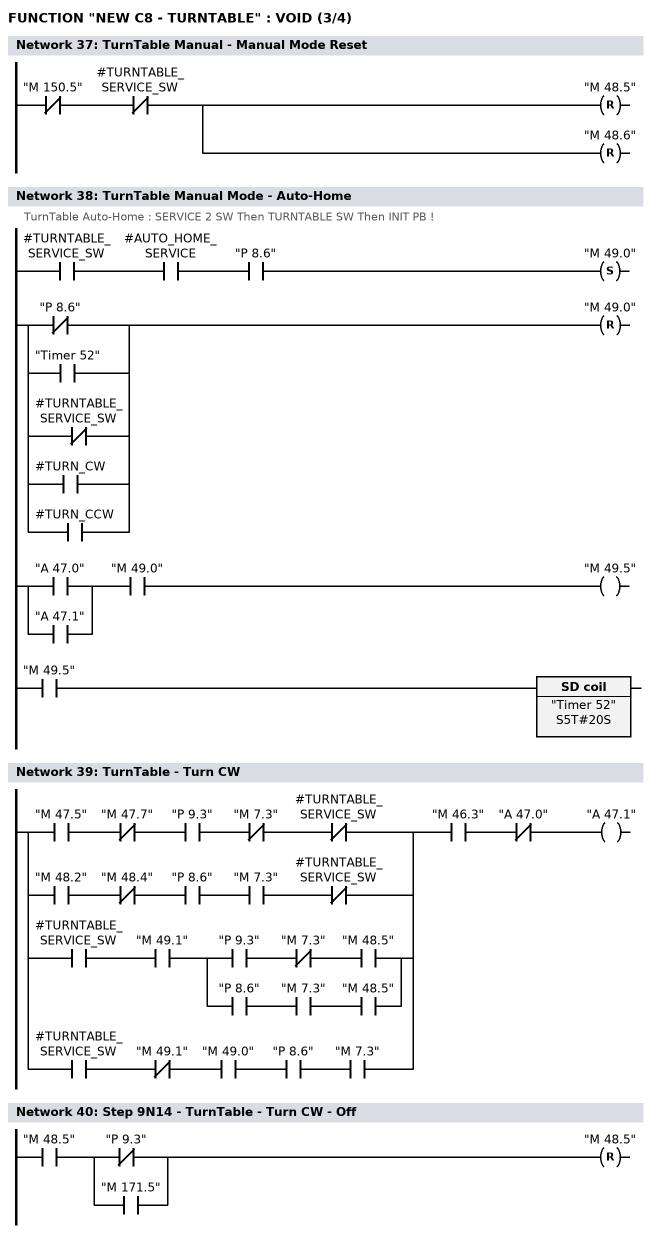

      AN    "M 150.5";
      AN    #TURNTABLE_SERVICE_SW;
      R     "M 48.5";
      R     "M 48.6";
NETWORK
TITLE =TurnTable Manual Mode - Auto-Home
//TurnTable Auto-Home : SERVICE 2 SW Then TURNTABLE SW Then INIT PB !
      A     #TURNTABLE_SERVICE_SW;
      A     #AUTO_HOME_SERVICE;
      A     "P 8.6";
      S     "M 49.0";
//;
      AN    "P 8.6";
      O     "Timer 52";
      ON    #TURNTABLE_SERVICE_SW;
      O     #TURN_CW;
      O     #TURN_CCW;
      R     "M 49.0";
//;
      A(    ;
      O     "A 47.0";
      O     "A 47.1";
      )     ;
      A     "M 49.0";
      =     "M 49.5";
//;
      A     "M 49.5";
      L     S5T#20S;
      SD    "Timer 52";
NETWORK
TITLE =TurnTable - Turn CW

      A(    ;
      A     "M 47.5";
      AN    "M 47.7";
      A     "P 9.3";
      AN    "M 7.3";
      AN    #TURNTABLE_SERVICE_SW;
      O     ;
      A     "M 48.2";
      AN    "M 48.4";
      A     "P 8.6";
      A     "M 7.3";
      AN    #TURNTABLE_SERVICE_SW;
      O     ;
      A     #TURNTABLE_SERVICE_SW;
      A     "M 49.1";
      A(    ;
      A     "P 9.3";
      AN    "M 7.3";
      A     "M 48.5";
      O     ;
      A     "P 8.6";
      A     "M 7.3";
      A     "M 48.5";
      )     ;
      O     ;
      A     #TURNTABLE_SERVICE_SW;
      AN    "M 49.1";
      A     "M 49.0";
      A     "P 8.6";
      A     "M 7.3";
      )     ;
      A     "M 46.3";
      AN    "A 47.0";
      =     "A 47.1";
NETWORK
TITLE =Step 9N14 - TurnTable - Turn CW - Off

      A     "M 48.5";
      A(    ;
      ON    "P 9.3";
      O     "M 171.5";
      )     ;
      R     "M 48.5";
NETWORK
TITLE =Turn Table - Turn CCW
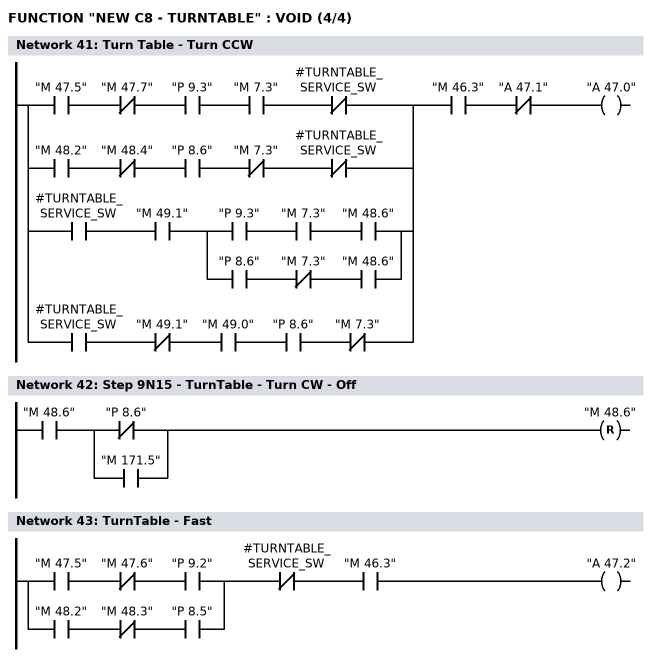

      A(    ;
      A     "M 47.5";
      AN    "M 47.7";
      A     "P 9.3";
      A     "M 7.3";
      AN    #TURNTABLE_SERVICE_SW;
      O     ;
      A     "M 48.2";
      AN    "M 48.4";
      A     "P 8.6";
      AN    "M 7.3";
      AN    #TURNTABLE_SERVICE_SW;
      O     ;
      A     #TURNTABLE_SERVICE_SW;
      A     "M 49.1";
      A(    ;
      A     "P 9.3";
      A     "M 7.3";
      A     "M 48.6";
      O     ;
      A     "P 8.6";
      AN    "M 7.3";
      A     "M 48.6";
      )     ;
      O     ;
      A     #TURNTABLE_SERVICE_SW;
      AN    "M 49.1";
      A     "M 49.0";
      A     "P 8.6";
      AN    "M 7.3";
      )     ;
      A     "M 46.3";
      AN    "A 47.1";
      =     "A 47.0";
NETWORK
TITLE =Step 9N15 - TurnTable - Turn CW - Off

      A     "M 48.6";
      A(    ;
      ON    "P 8.6";
      O     "M 171.5";
      )     ;
      R     "M 48.6";
NETWORK
TITLE =TurnTable - Fast

      A(    ;
      A     "M 47.5";
      AN    "M 47.6";
      A     "P 9.2";
      O     ;
      A     "M 48.2";
      AN    "M 48.3";
      A     "P 8.5";
      )     ;
      AN    #TURNTABLE_SERVICE_SW;
      A     "M 46.3";
      =     "A 47.2";
NETWORK
TITLE =TurnTable Position : Home = DB50.238:1 / Delivery = DB50.238:2

      OPN   "DB LAUER";
      ON    "P 8.6";
      ON    "P 9.3";
      JC    M003;
      L     W#16#0;
      T     DBW  238;
      BEC   ;

M003: A     "P 8.6";
      JC    M004;
      L     W#16#1;
      T     DBW  238;
      BEC   ;

M004: L     W#16#2;
      T     DBW  238;
END_FUNCTION

FUNCTION "NEW C9 - PUSHER 2" : VOID
TITLE =NEW FC950 (was FC1050) - Conveyor 9 / Pusher 2 Pos.11
//
//v1.0 2026-11-24: OMRON HMI positioning time (Timer 62) per packet length class
//from DB15 "PACKET POSITION DB".C9_Stop_S5T (FC1215 "PACKET POSITIONING", called
//by FC942). Class without time = "HMI_DB".CONV_9_POS_mS x 10 as before.
//v1.1 2026-11-24: DB15 symbol renamed "PACKET POSITION DB" - no code change.
NAME : POS_11
VERSION : 1.1


VAR_TEMP
  MAIN_SERVICE_2_SW : BOOL ;
  CONVEYOR_9_RUN : BOOL ;
  PUSHER_PUSH : BOOL ;
  INITIALISATION : BOOL ;
  POSITION_TIME : S5TIME ;
  ZOOLOO : TIME ;
END_VAR
BEGIN
NETWORK
TITLE =Pusher 2 - Service

      A     "HMI_DB".ALL_SERVICE_ENABLE_SW;
      A     "HMI_DB".CONVEYOR_9_SERVICE_SW;
      A     "HMI_DB".SERVICE_SW_2_STATUS;
      =     #MAIN_SERVICE_2_SW;
//;
      A     #MAIN_SERVICE_2_SW;
      O     "M 50.1";
      JNB   CON9;
      A     "HMI_DB".HMI_CONVEYOR_9_TEST_SSW;
      =     #CONVEYOR_9_RUN;
//;
      A     "HMI_DB".HMI_PUSHER_2_TEST_SSW;
      =     #PUSHER_PUSH;
//;
      A     "HMI_DB".SERVICE_INIT_PB;
      =     #INITIALISATION;
//;
      A     #CONVEYOR_9_RUN;
      S     "DB UTILITY".Conveyor_8_Disable;
//;
      A     #PUSHER_PUSH;
      S     "DB UTILITY".Conveyor_9_Disable;
//;
      AN    #MAIN_SERVICE_2_SW;
      R     "HMI_DB".HMI_CONVEYOR_9_TEST_SSW;
      R     "HMI_DB".HMI_PUSHER_2_TEST_SSW;
      R     "DB UTILITY".Conveyor_8_Disable;
      R     "DB UTILITY".Conveyor_9_Disable;

CON9: R     #CONVEYOR_9_RUN;
      R     #PUSHER_PUSH;
      R     #INITIALISATION;
      FP    "FP 169.1";
      =     "M 50.1";
NETWORK
TITLE =Pusher Rollers - Max Run Time

      A     "M 51.2";
      AN    "M 51.3";
      A     "M 0.3";
      L     S5T#5S;
      SD    "Timer 51";
NETWORK
TITLE =Conveyor 9 - Pusher Steps Register - Reset

      A(    ;
      A     "M 52.1";
      O     "Timer 51";
      O     #INITIALISATION;
      O     "DB UTILITY".Conveyor_9_Disable;
      )     ;
      A     "M 0.3";
      JC    M001;
      JU    M002;

M001: L     W#16#0;
      T     "MW 51";
      T     "MB 53";

M002: NOP   0;
NETWORK
TITLE =Step 10N1 - Power ON
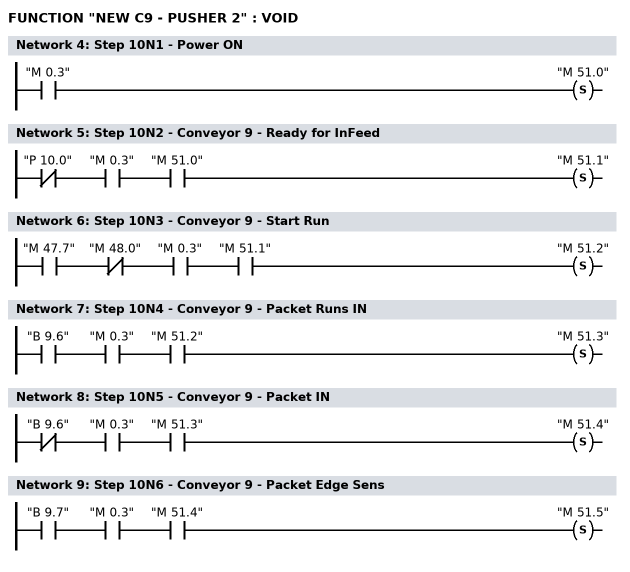

      A     "M 0.3";
      S     "M 51.0";
NETWORK
TITLE =Step 10N2 - Conveyor 9 - Ready for InFeed

      AN    "P 10.0";
      A     "M 0.3";
      A     "M 51.0";
      S     "M 51.1";
NETWORK
TITLE =Step 10N3 - Conveyor 9 - Start Run

      A     "M 47.7";
      AN    "M 48.0";
      A     "M 0.3";
      A     "M 51.1";
      S     "M 51.2";
NETWORK
TITLE =Step 10N4 - Conveyor 9 - Packet Runs IN

      A     "B 9.6";
      A     "M 0.3";
      A     "M 51.2";
      S     "M 51.3";
NETWORK
TITLE =Step 10N5 - Conveyor 9 - Packet IN

      AN    "B 9.6";
      A     "M 0.3";
      A     "M 51.3";
      S     "M 51.4";
NETWORK
TITLE =Step 10N6 - Conveyor 9 - Packet Edge Sens

      A     "B 9.7";
      A     "M 0.3";
      A     "M 51.4";
      S     "M 51.5";
NETWORK
TITLE =Time Convertion - Lateral Packet Position to Feeder - Adj.(HMI)

      A     "M 140.3";
      AN    "M 6.7";
      FP    "FP 147.2";
      JNB   BYP1;
      L     "HMI_DB".CONV_9_POS_mS; // Integer contains MILLISECOND seconds
      L     10;
      *I    ;
      ITD   ;
      T     #ZOOLOO;

      CALL "TIM_S5TI" (
           IN                       := #ZOOLOO,
           RET_VAL                  := #POSITION_TIME);

      L     #POSITION_TIME;
      T     "MW 184";
BYP1: CLR   ;

      A     "M 140.3";
      A     "M 51.5";
      AN    "M 51.6";
      A     "M 0.3";
      L     "PACKET POSITION DB".C9_Stop_S5T; // Was MW 184 - Now per Length Class (DB15)
      SD    "Timer 62"; // OMRON HMI
NETWORK
TITLE =Conveyor 9 - Lateral Packet Position to Feeder - Adj.(HMI)

      AN    "M 140.3";
      AN    "M 6.7";
      FP    "FP 149.5";
      JNB   BYP2;
      OPN   "DB LAUER";
      CALL "LAUER TIME" (
           QUEL                     := DBW  248,
           _TIME                    := MW   124);

BYP2: NOP   0;

      AN    "M 140.3";
      A     "M 51.5";
      AN    "M 51.6";
      A     "M 0.3";
      L     MW   124;
      SD    "Timer 50"; // LAUER HMI
NETWORK
TITLE =Step 10N7 - Conveyor 9 - Packet in Position - Stop
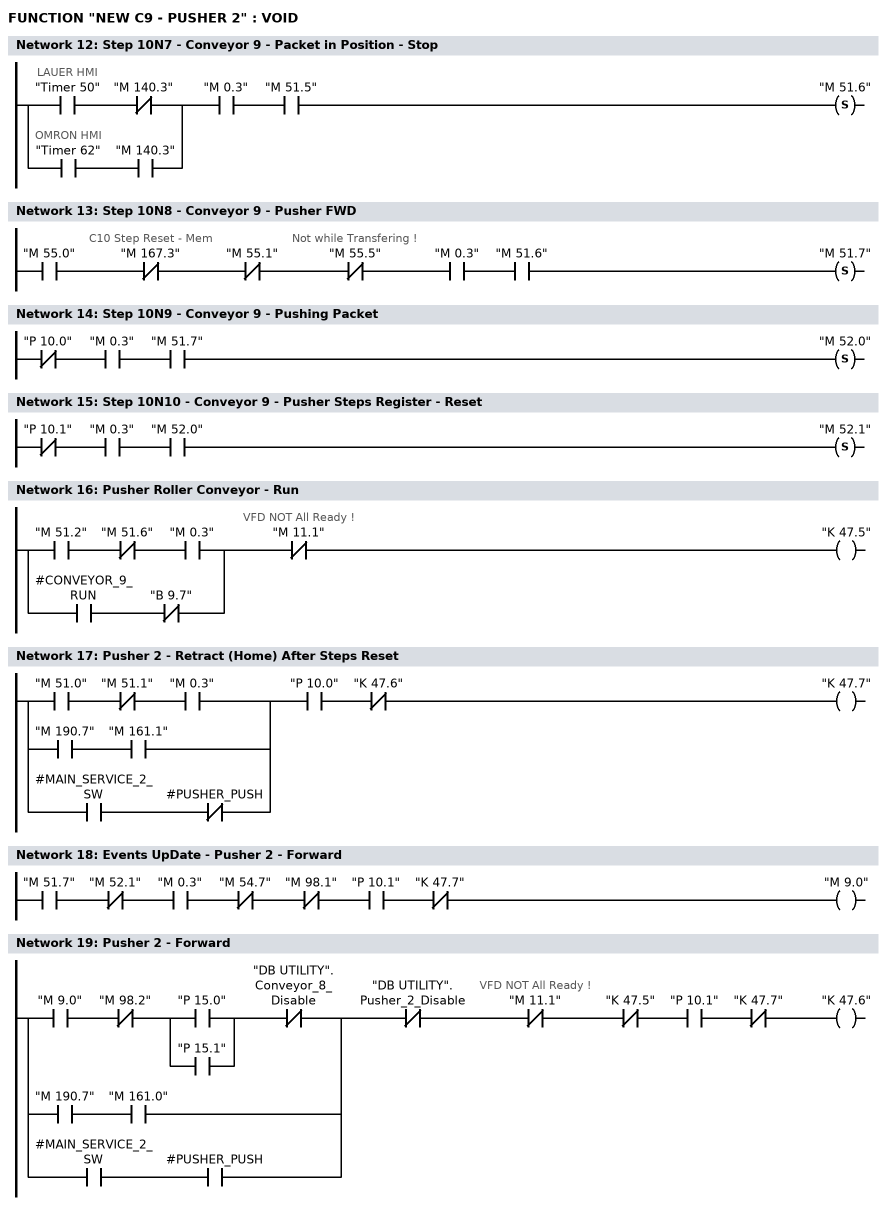

      A(    ;
      O(    ;
      A     "Timer 50"; // LAUER HMI
      AN    "M 140.3";
      )     ;
      O(    ;
      A     "Timer 62"; // OMRON HMI
      A     "M 140.3";
      )     ;
      )     ;
      A     "M 0.3";
      A     "M 51.5";
      S     "M 51.6";
NETWORK
TITLE =Step 10N8 - Conveyor 9 - Pusher FWD

      A     "M 55.0";
      AN    "M 167.3"; // C10 Step Reset - Mem
      AN    "M 55.1";
      AN    "M 55.5"; // Not while Transfering !
      A     "M 0.3";
      A     "M 51.6";
      S     "M 51.7";
NETWORK
TITLE =Step 10N9 - Conveyor 9 - Pushing Packet

      AN    "P 10.0";
      A     "M 0.3";
      A     "M 51.7";
      S     "M 52.0";
NETWORK
TITLE =Step 10N10 - Conveyor 9 - Pusher Steps Register - Reset

      AN    "P 10.1";
      A     "M 0.3";
      A     "M 52.0";
      S     "M 52.1";
NETWORK
TITLE =Pusher Roller Conveyor - Run

      A     "M 51.2";
      AN    "M 51.6";
      A     "M 0.3";
      O(    ;
      A     #CONVEYOR_9_RUN;
      AN    "B 9.7";
      )     ;
      AN    "M 11.1"; // VFD NOT All Ready !
      =     "K 47.5";
NETWORK
TITLE =Pusher 2 - Retract (Home) After Steps Reset

      A(    ;
      A     "M 51.0";
      AN    "M 51.1";
      A     "M 0.3";
      O     ;
      A     "M 190.7";
      A     "M 161.1";
      O     ;
      A     #MAIN_SERVICE_2_SW;
      AN    #PUSHER_PUSH;
      )     ;
      A     "P 10.0";
      AN    "K 47.6";
      =     "K 47.7";
NETWORK
TITLE =Events UpDate - Pusher 2 - Forward

      A     "M 51.7";
      AN    "M 52.1";
      A     "M 0.3";
      AN    "M 54.7";
      AN    "M 98.1";
      A     "P 10.1";
      AN    "K 47.7";
      =     "M 9.0";
NETWORK
TITLE =Pusher 2 - Forward

      A(    ;
      A     "M 9.0";
      AN    "M 98.2";
      A(    ;
      O     "P 15.0";
      O     "P 15.1";
      )     ;
      AN    "DB UTILITY".Conveyor_8_Disable;
      O     ;
      A     "M 190.7";
      A     "M 161.0";
      O     ;
      A     #MAIN_SERVICE_2_SW;
      A     #PUSHER_PUSH;
      )     ;
      AN    "DB UTILITY".Pusher_2_Disable;
      AN    "M 11.1"; // VFD NOT All Ready !
      AN    "K 47.5";
      A     "P 10.1";
      AN    "K 47.7";
      =     "K 47.6";
NETWORK
TITLE =Position Data Return

      OPN   "DB LAUER";
//;
      ON    "P 10.0";
      ON    "P 10.1";
      JC    M003;
      L     W#16#0;
      T     DBW  220;
      BEC   ;

M003: AN    "P 10.0";
      JC    M004;
      L     W#16#1;
      T     DBW  220;
      BEC   ;

M004: L     W#16#2;
      T     DBW  220;
END_FUNCTION

FUNCTION "NEW C10 - PIVOT PIW" : VOID
TITLE =FC 955 > NEW FC954 (was FC1054) - Pivot Conveyor 10 - Collator
//v0.1 2026-11-19: C10 encoder Ch5 read DIRECT every scan: PIW 334 (HW Config)
//instead
//of ACT_CNTV5. Ch4 (width gate) stays ACT_CNTV4: not in the direct area.
NAME : POS_12
VERSION : 0.1


VAR_TEMP
  MAIN_SERVICE_2_SW : BOOL ;
  PIVOT_SERVICE_SW : BOOL ;
  PIVOT_UP : BOOL ;
  PIVOT_DN : BOOL ;
  CONVEYOR_RUN : BOOL ;
  INITIALISATION : BOOL ;
  BARRIER_BLINKER : BOOL ;	//Feeder Safety Light Barrier
  PACKET_WIDTH_10 : WORD ;	//Collator Conveyor 10 - Packet Width
  FRAC_PACKET_WIDTH_10 : WORD ;	//Collator Conveyor 10 - Fraction of Packet Width
  PACKET_WIDTH_FRAC_10 : WORD ;	//Collator Conveyor 10 - Packet Width + Fraction
  SURFACE_LENGTH_LEFT_10 : WORD ;	//Collator Conveyor 10 - Surface Length Left
  QTY_MAX_10 : REAL ;
END_VAR
BEGIN
NETWORK
TITLE =Pivot Service

      A     "HMI_DB".ALL_SERVICE_ENABLE_SW;
      A     "HMI_DB".CONVEYOR_10_SERVICE_SW;
      A     "HMI_DB".SERVICE_SW_2_STATUS;
      =     #MAIN_SERVICE_2_SW;
//;
      A     #MAIN_SERVICE_2_SW;
      O     "M 54.3";
      JNB   PIVO;

      A     "HMI_DB".HMI_PIVOT_SERVICE_SSW;
      =     #PIVOT_SERVICE_SW;
      R     "HMI_DB".HMI_CONVEYOR_10_TEST_SSW;
//;
      A     "HMI_DB".HMI_CONVEYOR_10_TEST_SSW;
      =     #CONVEYOR_RUN;
      R     "HMI_DB".HMI_PIVOT_SERVICE_SSW;
//;
      A(    ;
      O     #PIVOT_SERVICE_SW;
      O     #CONVEYOR_RUN;
      )     ;
      S     "DB UTILITY".Pusher_2_Disable;
//;
      A     #PIVOT_SERVICE_SW;
      A     "HMI_DB".HMI_PIVOT_TEST_DN_SSW;
      AN    "HMI_DB".HMI_PIVOT_TEST_UP_SSW; // Not Both Switches
      =     #PIVOT_DN;
//;
      A     #PIVOT_SERVICE_SW;
      A     "HMI_DB".HMI_PIVOT_TEST_UP_SSW;
      AN    "HMI_DB".HMI_PIVOT_TEST_DN_SSW; // Not Both Switches
      =     #PIVOT_UP;
//;
      AN(   ;
      O     "P 15.0";
      O     "P 15.1";
      )     ;
      R     #CONVEYOR_RUN;
//;
      A     "HMI_DB".SERVICE_INIT_PB;
      =     #INITIALISATION;
//;
      AN    #MAIN_SERVICE_2_SW;
      R     "HMI_DB".HMI_PIVOT_SERVICE_SSW;
      R     "HMI_DB".HMI_CONVEYOR_10_TEST_SSW;
      R     "HMI_DB".HMI_PIVOT_TEST_DN_SSW;
      R     "HMI_DB".HMI_PIVOT_TEST_UP_SSW;
      R     "DB UTILITY".Pusher_2_Disable;

PIVO: R     #PIVOT_SERVICE_SW;
      R     #CONVEYOR_RUN;
      R     #INITIALISATION;
      R     #PIVOT_DN;
      R     #PIVOT_UP;
      FP    "FP 169.2";
      =     "M 54.3";
NETWORK
TITLE =Conveyor 10 - Packet Width - Measurements [mS]

      A     "B 10.4"; // C10 InFeed Sens
      A     "M 55.1"; // Collator Trigger - Step
      S     "M 166.4";
//;
      A     "M 166.4";
      =     "FM350 DB".CONTROL_SIGNALS.SW_GATE4;
//;
      A     "M 166.4";
      FP    "FP 149.7";
      JNB   NRAZ;
      L     0;
      T     "COLLATORS DB".Packet_Width_C10_mS;

NRAZ: A     "M 166.4";
      JNB   NCNT;
      L     "COLLATORS DB".Packet_Width_C10_mS;
      L     "DB UTILITY".Scan_Cycle_Previous;
      ITD   ;
      +D    ;
      T     "COLLATORS DB".Packet_Width_C10_mS;

NCNT: A     "M 166.4";
      AN    "B 10.4";
      JNB   M104;
      L     "FM350 DB".ACT_CNTV4; // C10 Encoder Counter
      T     #PACKET_WIDTH_10;
      T     "COLLATORS DB".Packet_Width_C10;
//;
      L     #PACKET_WIDTH_10;
      ITD   ;
      DTR   ;
      L     2.000000e-001;
      *R    ;
      RND   ;

      T     "COLLATORS DB".Frac_Packet_Width_C10;

      T     #FRAC_PACKET_WIDTH_10;
      L     #PACKET_WIDTH_10;
      +I    ;
      T     "COLLATORS DB".Packet_Width_Frac_C10;
      T     #PACKET_WIDTH_FRAC_10;
      R     "M 166.4";
      S     "M 167.2";

M104: NOP   0;
NETWORK
TITLE =Conveyor 10 - Packet Width Measurements [mm] - While Collating

      A     "B 10.4"; // C10 InFeed Sens - New Packet
      FP    "M 188.5";
      A     "A 48.0";
      JCN   NPRT;

      L     "PIW 334"; // Direct Ch5 (was ACT_CNTV5, ~100 mS old) C10 Encoder Counter
      T     "HOUSE_KEEPING DB".C10_Encoder_READ_Mem;

NPRT: AN    "B 10.4"; // C10 InFeed Sens - New Packet End
      FP    "M 188.6";
      JCN   NTKE;

      L     "PIW 334"; // Direct Ch5 (was ACT_CNTV5, ~100 mS old) C10 Encoder Counter
      L     "HOUSE_KEEPING DB".C10_Encoder_READ_Mem;
      -I    ;
      T     "HOUSE_KEEPING DB".C10_Packet_Width_ep; // C4 Packet Length [ep]
      DTR   ;
//;
      L     3.100000e-001; //  Encoder Wheel 283mm / 600 PPR  [mm/pulse]
      *R    ;
      RND   ;
      T     "HOUSE_KEEPING DB".C10_Packet_Width_mm;

NTKE: NOP   0;
NETWORK
TITLE =Conveyor 10 - Packet Width Measurements [mS]
//Conveyor 10 - Packet Width Measurements [mS]


NETWORK
TITLE =Conveyor 10 - Surface Length Left (PulseUnit) - Measurements

      A     "M 166.5";
      =     "FM350 DB".CONTROL_SIGNALS.SW_GATE5;
//;
      A     "M 166.5";
      JNB   M665;
      L     "COLLATORS DB".Surface_Length_10;
      L     "PIW 334"; // Direct Ch5 (was ACT_CNTV5, ~100 mS old)
      -D    ;
      T     #SURFACE_LENGTH_LEFT_10;
      L     0;
      >=I   ;
      JNB   T010;
      L     #SURFACE_LENGTH_LEFT_10;
      T     "COLLATORS DB".Surface_Length_Left_10;

T010: NOP   0;

M665: NOP   0;

      A     "M 55.1"; // Collator Trigger
      FP    "FP 154.6";
      S     "M 166.5";
NETWORK
TITLE =Conveyor 10 - Space Between Packet - Calculator
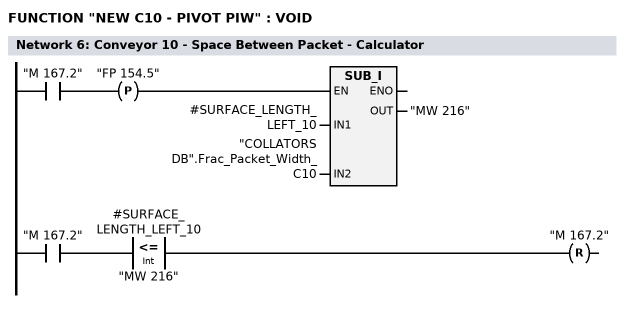

      A     "M 167.2";
      FP    "FP 154.5";
      JNB   M582;
      L     #SURFACE_LENGTH_LEFT_10;
      L     "COLLATORS DB".Frac_Packet_Width_C10;
      -I    ;
      T     "MW 216";

M582: NOP   0;

      A     "M 167.2";
      A(    ;
      L     #SURFACE_LENGTH_LEFT_10;
      L     "MW 216";
      <=I   ;
      )     ;
      R     "M 167.2";
NETWORK
TITLE =Conveyor 10 - Collating Surface Manager

      A     "M 166.5";
      AN    "M 55.4";
      AN    "M 54.4"; // Collator Full - Count Flag Off
      A     "M 55.3";
      JNB   M554;

      A(    ;
      L     #SURFACE_LENGTH_LEFT_10;
      L     "COLLATORS DB".Packet_Width_Frac_C10;
      <I    ;
      )     ;
      S     "M 54.4"; // Collator Full - Count - Set

M554: NOP   0;

      A     "M 167.3"; // C10 Step Reset - Mem
      R     "M 54.4"; // Collator Full - Count - Reset
NETWORK
TITLE =Conveyor 10 - Surface Length Reset

      ON(   ;
      O     "P 15.0"; // While C10 Pivoting...
      O     "P 15.1";
      )     ;
      L     S5T#200MS;
      SD    "Timer 104";
//;
      A     "Timer 104"; // C10 Surface Length Reset
      R     "M 166.4";
      R     "M 166.5";
NETWORK
TITLE =Clearing - C10 Counters Reset
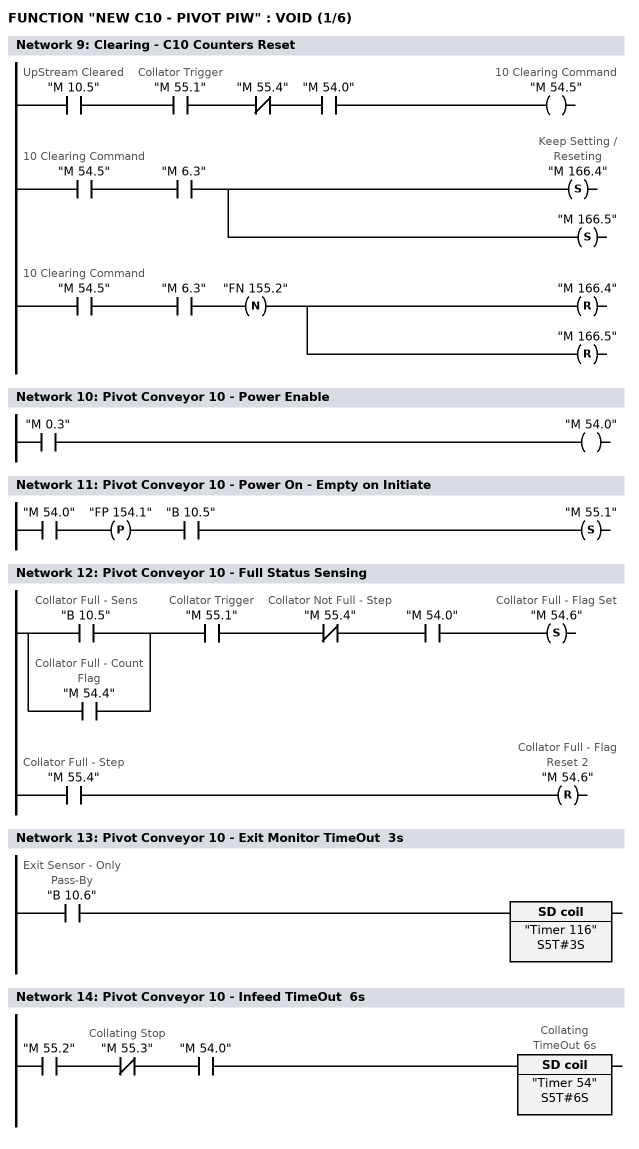

      A     "M 10.5"; // UpStream Cleared
      A     "M 55.1"; // Collator Trigger
      AN    "M 55.4";
      A     "M 54.0";
      =     "M 54.5"; // 10 Clearing Command
//;
      A     "M 54.5"; // 10 Clearing Command
      A     "M 6.3";
      S     "M 166.4"; // Keep Setting / Reseting
      S     "M 166.5";
//;
      A     "M 54.5"; // 10 Clearing Command
      A     "M 6.3";
      FN    "FN 155.2";
      R     "M 166.4";
      R     "M 166.5";
NETWORK
TITLE =Pivot Conveyor 10 - Power Enable

      A     "M 0.3";
      =     "M 54.0";
NETWORK
TITLE =Pivot Conveyor 10 - Power On - Empty on Initiate

      A     "M 54.0";
      FP    "FP 154.1"; // Empty on Power ON
      A     "B 10.5";
      S     "M 55.1";
NETWORK
TITLE =Pivot Conveyor 10 - Full Status Sensing

      A(    ;
      O     "B 10.5"; // Collator Full - Sens
      O     "M 54.4"; // Collator Full - Count Flag
      )     ;
      A     "M 55.1"; // Collator Trigger
      AN    "M 55.4"; // Collator Not Full - Step
      A     "M 54.0";
      S     "M 54.6"; // Collator Full - Flag Set
//;
      A     "M 55.4"; // Collator Full - Step
      R     "M 54.6"; // Collator Full - Flag Reset 2
NETWORK
TITLE =Pivot Conveyor 10 - Exit Monitor TimeOut  3s

      A     "B 10.6"; // Exit Sensor - Only Pass-By
      L     S5T#3S;
      SD    "Timer 116"; // Packet is Stuck !
NETWORK
TITLE =Pivot Conveyor 10 - Infeed TimeOut  6s

      A     "M 55.2";
      AN    "M 55.3"; // Collating Stop
      A     "M 54.0";
      L     S5T#6S; // Collating TimeOut 6s
      SD    "Timer 54";
NETWORK
TITLE =Pivot Conveyor 10 - Fault
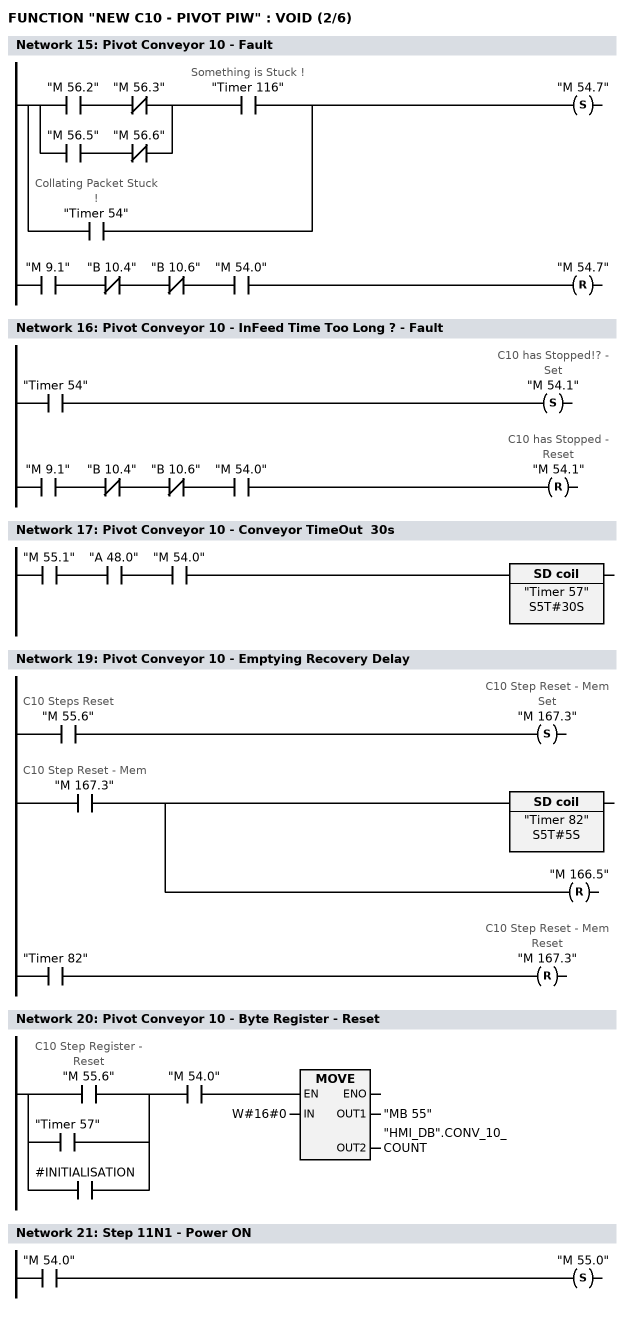

      A(    ;
      A(    ;
      A     "M 56.2";
      AN    "M 56.3";
      O     ;
      A     "M 56.5";
      AN    "M 56.6";
      )     ;
      A     "Timer 116"; // Something is Stuck !
      O     "Timer 54"; // Collating Packet Stuck !
      )     ;
      S     "M 54.7";
//;
      A     "M 9.1";
      AN    "B 10.4";
      AN    "B 10.6";
      A     "M 54.0";
      R     "M 54.7";
NETWORK
TITLE =Pivot Conveyor 10 - InFeed Time Too Long ? - Fault

      A     "Timer 54";
      S     "M 54.1"; // C10 has Stopped!? - Set
//;
      A     "M 9.1";
      AN    "B 10.4";
      AN    "B 10.6";
      A     "M 54.0";
      R     "M 54.1"; // C10 has Stopped - Reset
NETWORK
TITLE =Pivot Conveyor 10 - Conveyor TimeOut  30s

      A     "M 55.1";
      A     "A 48.0";
      A     "M 54.0";
      L     S5T#30S;
      SD    "Timer 57";
NETWORK
TITLE =Collating
//Collating


NETWORK
TITLE =Pivot Conveyor 10 - Emptying Recovery Delay

      A     "M 55.6"; // C10 Steps Reset
      S     "M 167.3"; // C10 Step Reset - Mem Set
//;
      A     "M 167.3"; // C10 Step Reset - Mem
      L     S5T#5S;
      SD    "Timer 82";
      R     "M 166.5";
//;
      A     "Timer 82";
      R     "M 167.3"; // C10 Step Reset - Mem Reset
NETWORK
TITLE =Pivot Conveyor 10 - Byte Register - Reset

      A(    ;
      O     "M 55.6"; // C10 Step Register - Reset
      O     "Timer 57";
      O     #INITIALISATION;
      )     ;
      A     "M 54.0";
      JNB   M001;
      L     W#16#0;
      T     "MB 55";
      T     "HMI_DB".CONV_10_COUNT;

M001: NOP   0;
NETWORK
TITLE =Step 11N1 - Power ON

      A     "M 54.0";
      S     "M 55.0";
NETWORK
TITLE =Step 11N2 - Conveyor 10 - Run
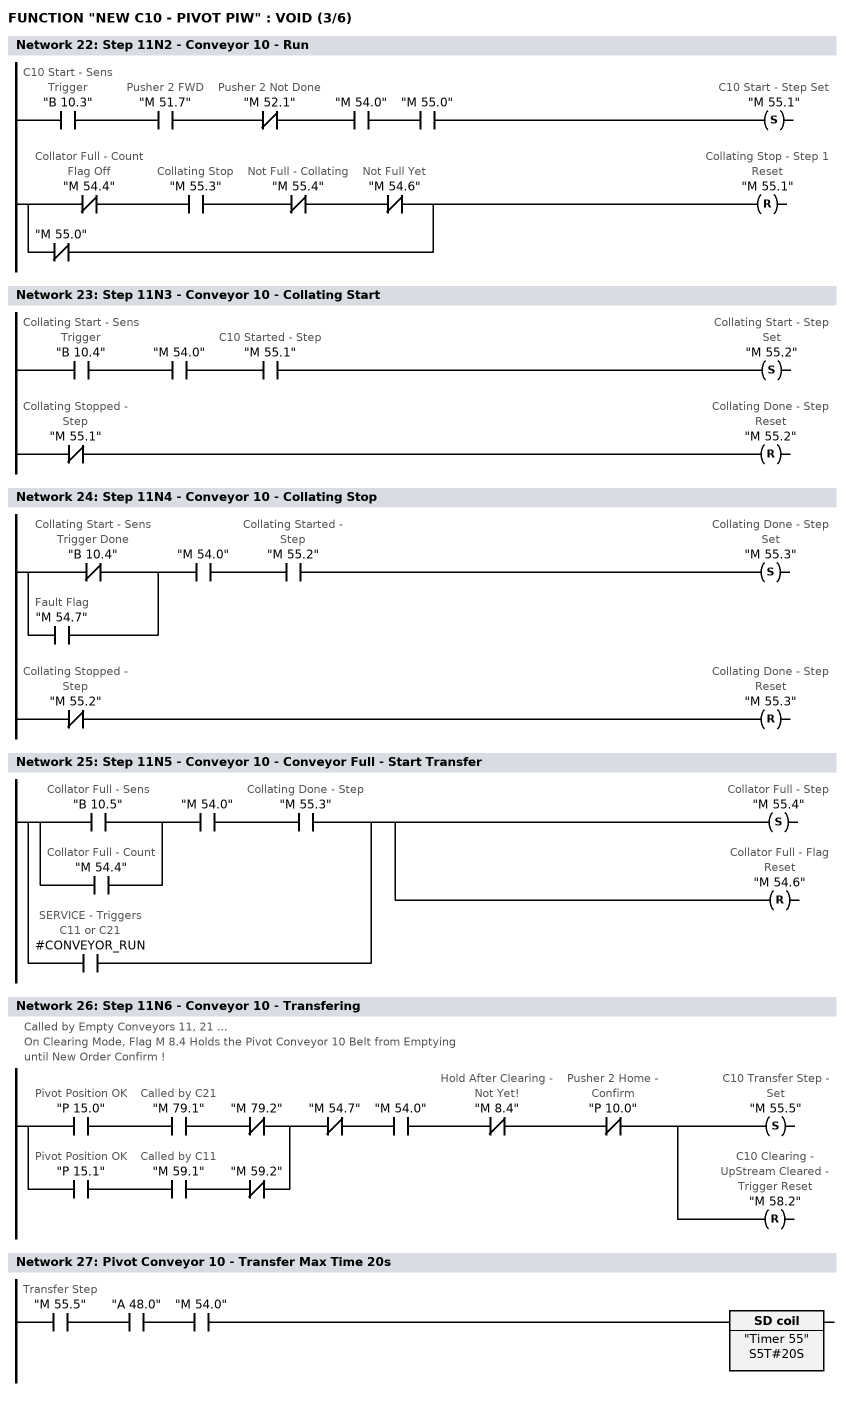

      A     "B 10.3"; // C10 Start - Sens Trigger
      A     "M 51.7"; // Pusher 2 FWD
      AN    "M 52.1"; // Pusher 2 Not Done
      A     "M 54.0";
      A     "M 55.0";
      S     "M 55.1"; // C10 Start - Step Set
//;
      A(    ;
      AN    "M 54.4"; // Collator Full - Count Flag Off
      A     "M 55.3"; // Collating Stop
      AN    "M 55.4"; // Not Full - Collating
      AN    "M 54.6"; // Not Full Yet
      ON    "M 55.0";
      )     ;
      R     "M 55.1"; // Collating Stop - Step 1 Reset
NETWORK
TITLE =Step 11N3 - Conveyor 10 - Collating Start

      A     "B 10.4"; // Collating Start - Sens Trigger
      A     "M 54.0";
      A     "M 55.1"; // C10 Started - Step
      S     "M 55.2"; // Collating Start - Step Set
//;
      AN    "M 55.1"; // Collating Stopped - Step
      R     "M 55.2"; // Collating Done - Step Reset
NETWORK
TITLE =Step 11N4 - Conveyor 10 - Collating Stop

      A(    ;
      ON    "B 10.4"; // Collating Start - Sens Trigger Done
      O     "M 54.7"; // Fault Flag
      )     ;
      A     "M 54.0";
      A     "M 55.2"; // Collating Started - Step
      S     "M 55.3"; // Collating Done - Step Set
//;
      AN    "M 55.2"; // Collating Stopped - Step
      R     "M 55.3"; // Collating Done - Step Reset
NETWORK
TITLE =Step 11N5 - Conveyor 10 - Conveyor Full - Start Transfer

      A(    ;
      O     "B 10.5"; // Collator Full - Sens
      O     "M 54.4"; // Collator Full - Count
      )     ;
      A     "M 54.0";
      A     "M 55.3"; // Collating Done - Step
      O     #CONVEYOR_RUN; // SERVICE - Triggers C11 or C21
      S     "M 55.4"; // Collator Full - Step
      R     "M 54.6"; // Collator Full - Flag Reset
NETWORK
TITLE =Step 11N6 - Conveyor 10 - Transfering
//Called by Empty Conveyors 11, 21 ...
//On Clearing Mode, Flag M 8.4 Holds the Pivot Conveyor 10 Belt from Emptying
//until New Order Confirm !
      A(    ;
      A     "P 15.0"; // Pivot Position OK
      A     "M 79.1"; // Called by C21
      AN    "M 79.2";
      O     ;
      A     "P 15.1"; // Pivot Position OK
      A     "M 59.1"; // Called by C11
      AN    "M 59.2";
      )     ;
      AN    "M 54.7";
      A     "M 54.0";
      AN    "M 8.4"; // Hold After Clearing - Not Yet!
      AN    "P 10.0"; // Pusher 2 Home - Confirm
      S     "M 55.5"; // C10 Transfer Step - Set
      R     "M 58.2"; // C10 Clearing - UpStream Cleared - Trigger Reset
NETWORK
TITLE =Pivot Conveyor 10 - Transfer Max Time 20s

      A     "M 55.5"; // Transfer Step
      A     "A 48.0";
      A     "M 54.0";
      L     S5T#20S;
      SD    "Timer 55"; // Transfer TimeOut
NETWORK
TITLE =Step 11N7 - Conveyor 10 - Steps Register - Reset
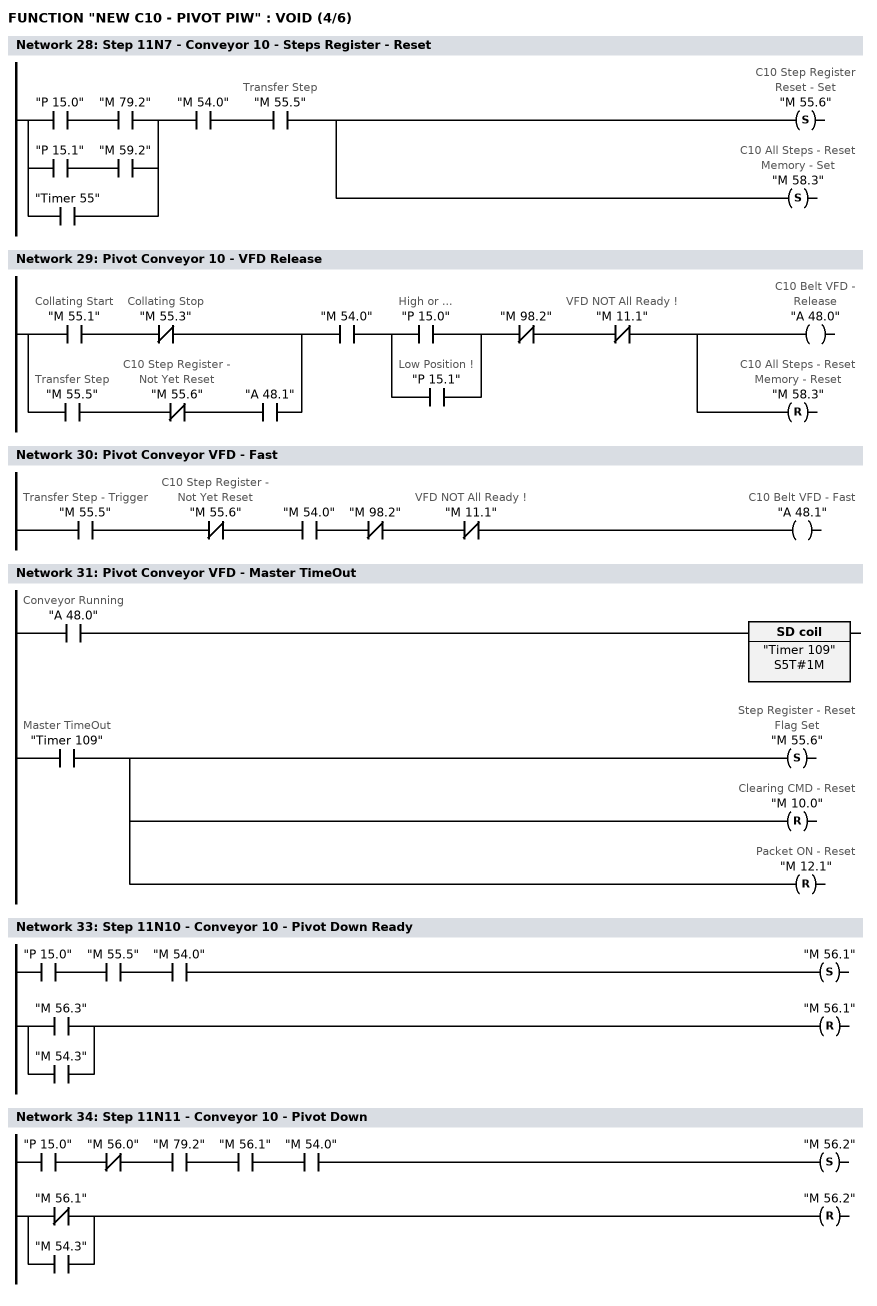

      A(    ;
      A     "P 15.0";
      A     "M 79.2";
      O     ;
      A     "P 15.1";
      A     "M 59.2";
      O     "Timer 55";
      )     ;
      A     "M 54.0";
      A     "M 55.5"; // Transfer Step
      S     "M 55.6"; // C10 Step Register Reset - Set
      S     "M 58.3"; // C10 All Steps - Reset Memory - Set
NETWORK
TITLE =Pivot Conveyor 10 - VFD Release

      A(    ;
      A     "M 55.1"; // Collating Start
      AN    "M 55.3"; // Collating Stop
      O     ;
      A     "M 55.5"; // Transfer Step
      AN    "M 55.6"; // C10 Step Register - Not Yet Reset
      A     "A 48.1";
      )     ;
      A     "M 54.0";
      A(    ;
      O     "P 15.0"; // High or ...
      O     "P 15.1"; // Low Position !
      )     ;
      AN    "M 98.2";
      AN    "M 11.1"; // VFD NOT All Ready !
      =     "A 48.0"; // C10 Belt VFD - Release
      R     "M 58.3"; // C10 All Steps - Reset Memory - Reset
NETWORK
TITLE =Pivot Conveyor VFD - Fast

      A     "M 55.5"; // Transfer Step - Trigger
      AN    "M 55.6"; // C10 Step Register - Not Yet Reset
      A     "M 54.0";
      AN    "M 98.2";
      AN    "M 11.1"; // VFD NOT All Ready !
      =     "A 48.1"; // C10 Belt VFD - Fast
NETWORK
TITLE =Pivot Conveyor VFD - Master TimeOut

      A     "A 48.0"; // Conveyor Running
      L     S5T#1M;
      SD    "Timer 109"; // Master TimeOut
//;
      A     "Timer 109"; // Master TimeOut
      S     "M 55.6"; // Step Register - Reset Flag Set
      R     "M 10.0"; // Clearing CMD - Reset
      R     "M 12.1"; // Packet ON - Reset
NETWORK
TITLE =Pivot Action
//Pivot Action


NETWORK
TITLE =Step 11N10 - Conveyor 10 - Pivot Down Ready

      A     "P 15.0";
      A     "M 55.5";
      A     "M 54.0";
      S     "M 56.1";
//;
      A     "M 56.3";
      O     "M 54.3";
      R     "M 56.1";
NETWORK
TITLE =Step 11N11 - Conveyor 10 - Pivot Down

      A     "P 15.0";
      AN    "M 56.0";
      A     "M 79.2";
      A     "M 56.1";
      A     "M 54.0";
      S     "M 56.2";
//;
      AN    "M 56.1";
      O     "M 54.3";
      R     "M 56.2";
NETWORK
TITLE =Step 11N12 - Conveyor 10 - Move Dn Stop
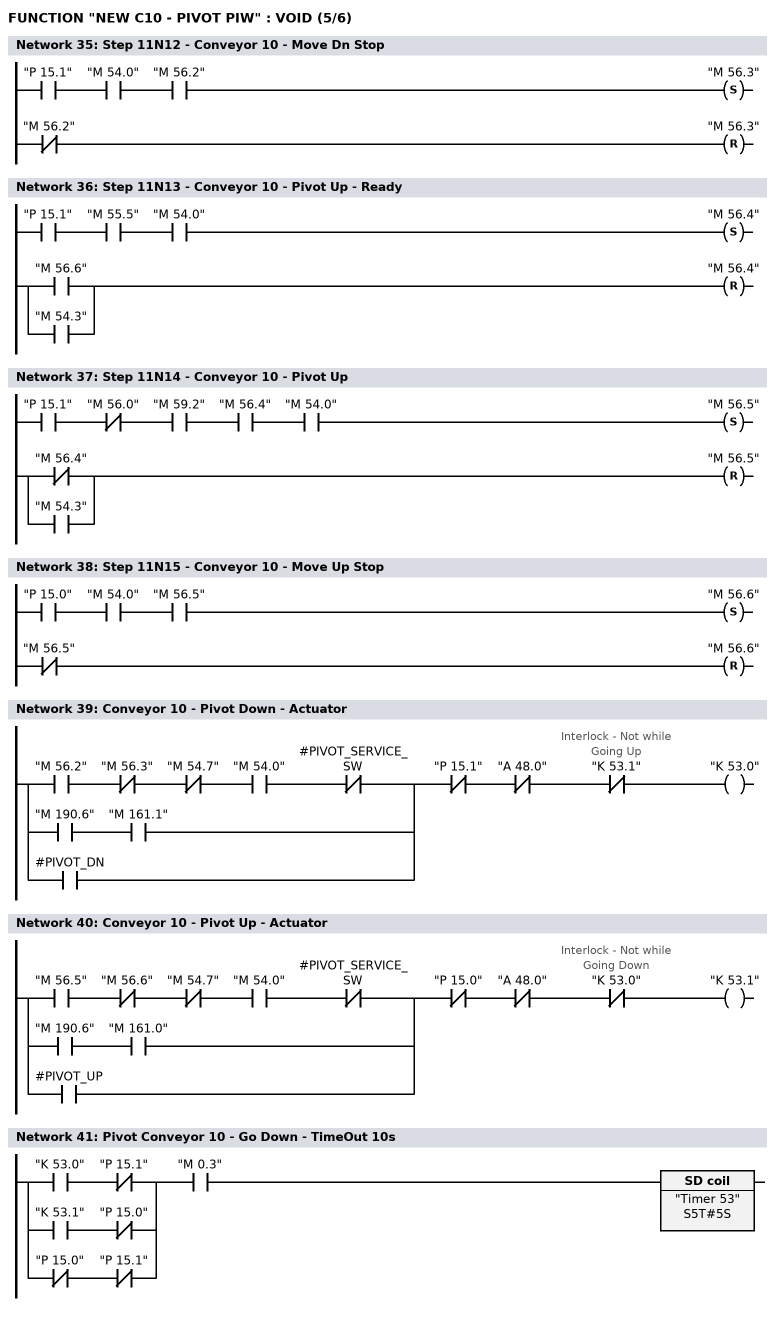

      A     "P 15.1";
      A     "M 54.0";
      A     "M 56.2";
      S     "M 56.3";
//;
      AN    "M 56.2";
      R     "M 56.3";
NETWORK
TITLE =Step 11N13 - Conveyor 10 - Pivot Up - Ready

      A     "P 15.1";
      A     "M 55.5";
      A     "M 54.0";
      S     "M 56.4";
//;
      A     "M 56.6";
      O     "M 54.3";
      R     "M 56.4";
NETWORK
TITLE =Step 11N14 - Conveyor 10 - Pivot Up

      A     "P 15.1";
      AN    "M 56.0";
      A     "M 59.2";
      A     "M 56.4";
      A     "M 54.0";
      S     "M 56.5";
//;
      AN    "M 56.4";
      O     "M 54.3";
      R     "M 56.5";
NETWORK
TITLE =Step 11N15 - Conveyor 10 - Move Up Stop

      A     "P 15.0";
      A     "M 54.0";
      A     "M 56.5";
      S     "M 56.6";
//;
      AN    "M 56.5";
      R     "M 56.6";
NETWORK
TITLE =Conveyor 10 - Pivot Down - Actuator

      A(    ;
      A     "M 56.2";
      AN    "M 56.3";
      AN    "M 54.7";
      A     "M 54.0";
      AN    #PIVOT_SERVICE_SW;
      O     ;
      A     "M 190.6";
      A     "M 161.1";
      )     ;
      O     #PIVOT_DN;
      AN    "P 15.1";
      AN    "A 48.0";
      AN    "K 53.1"; // Interlock - Not while Going Up
      =     "K 53.0";
NETWORK
TITLE =Conveyor 10 - Pivot Up - Actuator

      A(    ;
      A     "M 56.5";
      AN    "M 56.6";
      AN    "M 54.7";
      A     "M 54.0";
      AN    #PIVOT_SERVICE_SW;
      O     ;
      A     "M 190.6";
      A     "M 161.0";
      )     ;
      O     #PIVOT_UP;
      AN    "P 15.0";
      AN    "A 48.0";
      AN    "K 53.0"; // Interlock - Not while Going Down
      =     "K 53.1";
NETWORK
TITLE =Pivot Conveyor 10 - Go Down - TimeOut 10s

      A(    ;
      A     "K 53.0";
      AN    "P 15.1";
      O     ;
      A     "K 53.1";
      AN    "P 15.0";
      O     ;
      AN    "P 15.0";
      AN    "P 15.1";
      )     ;
      A     "M 0.3";
      L     S5T#5S;
      SD    "Timer 53";
NETWORK
TITLE =Pivot Conveyor 10 - Pivot Alarm
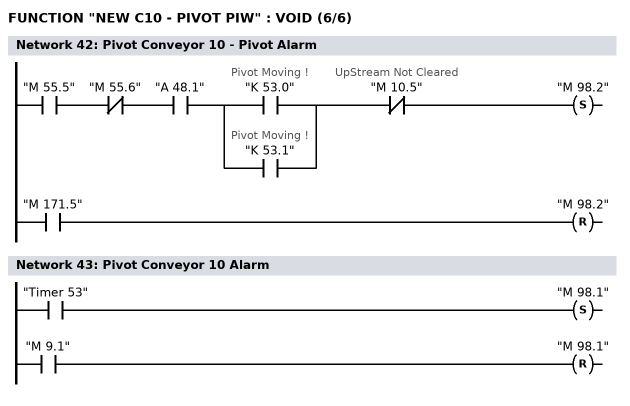

      A(    ;
      A     "M 55.5";
      AN    "M 55.6";
      A     "A 48.1";
      )     ;
      A(    ;
      O     "K 53.0"; // Pivot Moving !
      O     "K 53.1"; // Pivot Moving !
      )     ;
      AN    "M 10.5"; // UpStream Not Cleared
      S     "M 98.2";
//;
      A     "M 171.5";
      R     "M 98.2";
NETWORK
TITLE =Pivot Conveyor 10 Alarm

      A     "Timer 53";
      S     "M 98.1";
//;
      A     "M 9.1";
      R     "M 98.1";
NETWORK
TITLE =DBW  236 - Conveyor 10 - Position Transfer

      OPN   "DB LAUER";

      O     "P 15.0";
      O     "P 15.1";
      JC    M003;
      L     W#16#0;
      T     DBW  236;
      BEC   ;

M003: AN    "P 15.1";
      JC    M004;
      L     W#16#1;
      T     DBW  236;
      BEC   ;

M004: L     W#16#2;
      T     DBW  236;
END_FUNCTION

FUNCTION "NEW C11 - LINK 1 LO" : VOID
TITLE =NEW FC958 (was FC1058) - Conveyor 11 - Link 1L Pos. 13 Low Level
//
//v0.1 2026-11-19: clearing trigger M9.3 only if pivot LOW (P15.1).
NAME : POS_13_L
VERSION : 0.1


VAR_TEMP
  MAIN_SERVICE_2_SW : BOOL ;
  SERVICE_RUN : BOOL ;
  INITIALISATION : BOOL ;
  BARRIER_BLINKER : BOOL ;
END_VAR
BEGIN
NETWORK
TITLE =Conveyor 11 - Service

      A     "HMI_DB".ALL_SERVICE_ENABLE_SW;
      A     "HMI_DB".CONVEYOR_11_SERVICE_SW;
      A     "HMI_DB".SERVICE_SW_2_STATUS;
      =     #MAIN_SERVICE_2_SW;
//;
      A     #MAIN_SERVICE_2_SW;
      O     "M 58.7";
      JNB   CO11;
//;
      A     "HMI_DB".HMI_CONVEYOR_11_TEST_SSW;
      AN    "A 48.0";
      =     #SERVICE_RUN;
      S     "DB UTILITY".Conveyor_10_Disable;
      S     "DB UTILITY".Pivot_Disable;
//;
      A     "HMI_DB".SERVICE_INIT_PB;
      =     #INITIALISATION;
//;
      AN    #MAIN_SERVICE_2_SW;
      R     "HMI_DB".HMI_CONVEYOR_11_TEST_SSW;
      R     "DB UTILITY".Conveyor_10_Disable;
      R     "DB UTILITY".Pivot_Disable;

CO11: R     #SERVICE_RUN;
      R     #INITIALISATION;
      FP    "FP 148.0";
      =     "M 58.7";
NETWORK
TITLE =Power Enable
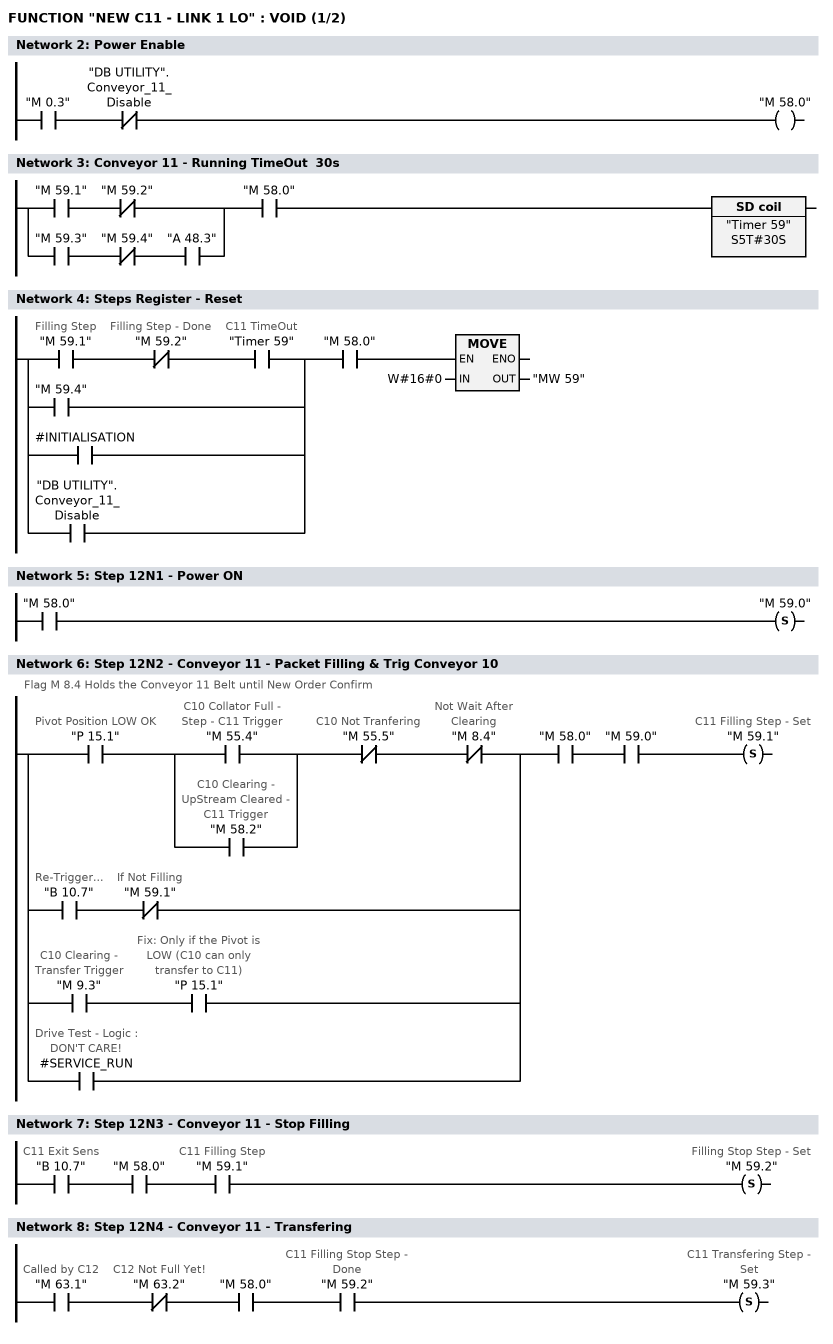

      A     "M 0.3";
      AN    "DB UTILITY".Conveyor_11_Disable;
      =     "M 58.0";
NETWORK
TITLE =Conveyor 11 - Running TimeOut  30s

      A(    ;
      A     "M 59.1";
      AN    "M 59.2";
      O     ;
      A     "M 59.3";
      AN    "M 59.4";
      A     "A 48.3";
      )     ;
      A     "M 58.0";
      L     S5T#30S;
      SD    "Timer 59"; // C11 TimeOut
NETWORK
TITLE =Steps Register - Reset

      A(    ;
      A     "M 59.1"; // Filling Step
      AN    "M 59.2"; // Filling Step - Done
      A     "Timer 59"; // C11 TimeOut
      O     "M 59.4";
      O     #INITIALISATION;
      O     "DB UTILITY".Conveyor_11_Disable;
      )     ;
      A     "M 58.0";
      JNB   _001;
      L     W#16#0;
      T     "MW 59";

_001: NOP   0;
NETWORK
TITLE =Step 12N1 - Power ON

      A     "M 58.0";
      S     "M 59.0";
NETWORK
TITLE =Step 12N2 - Conveyor 11 - Packet Filling & Trig Conveyor 10
//Flag M 8.4 Holds the Conveyor 11 Belt until New Order Confirm
      A(    ;
      A     "P 15.1"; // Pivot Position LOW OK
      A(    ;
      O     "M 55.4"; // C10 Collator Full - Step - C11 Trigger
      O     "M 58.2"; // C10 Clearing - UpStream Cleared - C11 Trigger
      )     ;
      AN    "M 55.5"; // C10 Not Tranfering
      AN    "M 8.4"; // Not Wait After Clearing
      O     ;
      A     "B 10.7"; // Re-Trigger...
      AN    "M 59.1"; // If Not Filling
      O     ;
      A     "M 9.3"; // C10 Clearing - Transfer Trigger
      A     "P 15.1"; // Fix: Only if the Pivot is LOW (C10 can only transfer to C11)
      )     ;
      O     #SERVICE_RUN; // Drive Test - Logic : DON'T CARE!
      A     "M 58.0";
      A     "M 59.0";
      S     "M 59.1"; // C11 Filling Step - Set
NETWORK
TITLE =Step 12N3 - Conveyor 11 - Stop Filling

      A     "B 10.7"; // C11 Exit Sens
      A     "M 58.0";
      A     "M 59.1"; // C11 Filling Step
      S     "M 59.2"; // Filling Stop Step - Set
NETWORK
TITLE =Step 12N4 - Conveyor 11 - Transfering

      A     "M 63.1"; // Called by C12
      AN    "M 63.2"; // C12 Not Full Yet!
      A     "M 58.0";
      A     "M 59.2"; // C11 Filling Stop Step - Done
      S     "M 59.3"; // C11 Transfering Step - Set
NETWORK
TITLE =Step 12N5 - Conveyor 11 - Steps Register - Reset
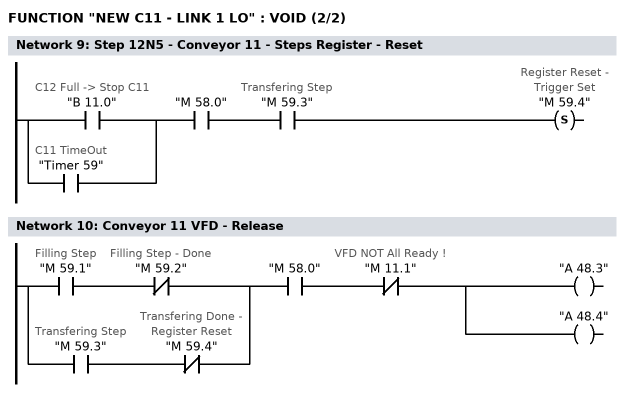

      A(    ;
      O     "B 11.0"; // C12 Full -> Stop C11
      O     "Timer 59"; // C11 TimeOut
      )     ;
      A     "M 58.0";
      A     "M 59.3"; // Transfering Step
      S     "M 59.4"; // Register Reset - Trigger Set
NETWORK
TITLE =Conveyor 11 VFD - Release

      A(    ;
      A     "M 59.1"; // Filling Step
      AN    "M 59.2"; // Filling Step - Done
      O     ;
      A     "M 59.3"; // Transfering Step
      AN    "M 59.4"; // Transfering Done - Register Reset
      )     ;
      A     "M 58.0";
      AN    "M 11.1"; // VFD NOT All Ready !
      =     "A 48.3";
      =     "A 48.4";
END_FUNCTION

FUNCTION "NEW C12 - LINK 2 LO" : VOID
TITLE =NEW FC962 (was FC1062) - Conveyor 12 - Link 2L Pos. 14 Low Level
//
NAME : POS_14_L
VERSION : 0.0


VAR_TEMP
  MAIN_SERVICE_2_SW : BOOL ;
  SERVICE_RUN : BOOL ;
  BARRIER_BLINKER : BOOL ;
END_VAR
BEGIN
NETWORK
TITLE =Conveyor 12 - Service

      A     "HMI_DB".ALL_SERVICE_ENABLE_SW;
      A     "HMI_DB".CONVEYOR_11_SERVICE_SW;
      A     "HMI_DB".SERVICE_SW_2_STATUS;
      =     #MAIN_SERVICE_2_SW;
//;
      A     #MAIN_SERVICE_2_SW;
      O     "M 62.7";
      JNB   CO12;
//;
      A     "HMI_DB".HMI_CONVEYOR_12_TEST_SSW;
      =     #SERVICE_RUN;
//;
      AN    #MAIN_SERVICE_2_SW;
      R     "HMI_DB".HMI_CONVEYOR_12_TEST_SSW;

CO12: R     #SERVICE_RUN;
      FP    "FP 148.1";
      =     "M 62.7";
NETWORK
TITLE =FL Power Enable
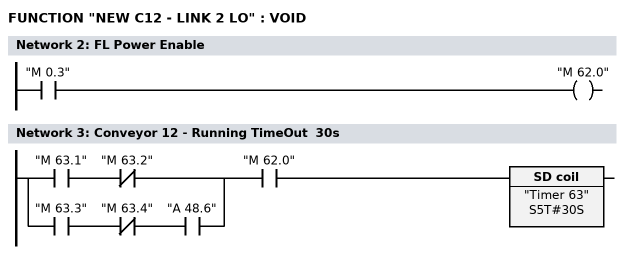

      A     "M 0.3";
      =     "M 62.0";
NETWORK
TITLE =Conveyor 12 - Running TimeOut  30s

      A(    ;
      A     "M 63.1";
      AN    "M 63.2";
      O     ;
      A     "M 63.3";
      AN    "M 63.4";
      A     "A 48.6";
      )     ;
      A     "M 62.0";
      L     S5T#30S;
      SD    "Timer 63";
NETWORK
TITLE =Conveyor 12 - Steps Register - Reset

      A(    ;
      A     "M 63.1";
      AN    "M 63.2";
      A     "Timer 63";
      O     "M 63.4";
      )     ;
      A     "M 62.0";
      JC    M001;
      JU    M002;

M001: L     W#16#0;
      T     "MW 63";
      T     "MB 65";

M002: NOP   0;
NETWORK
TITLE =Step 13N1 - Power On
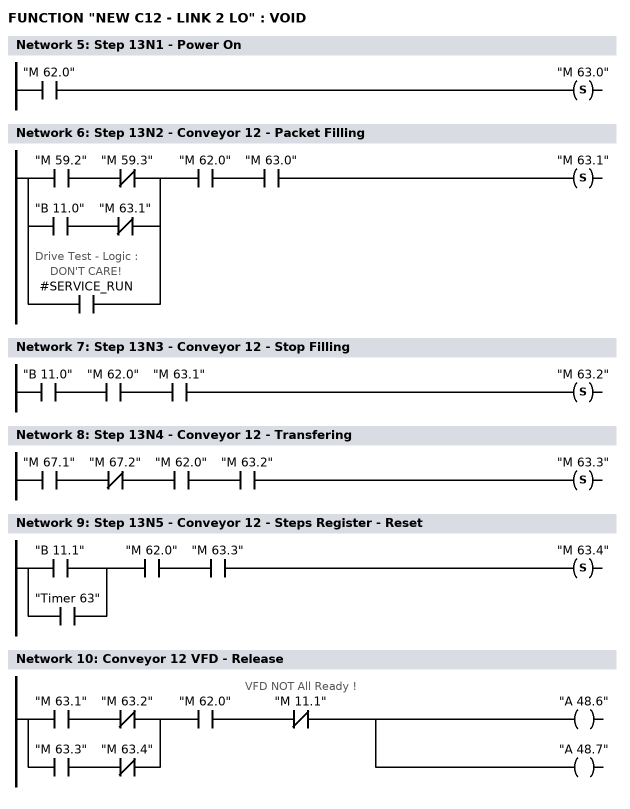

      A     "M 62.0";
      S     "M 63.0";
NETWORK
TITLE =Step 13N2 - Conveyor 12 - Packet Filling

      A(    ;
      A     "M 59.2";
      AN    "M 59.3";
      O     ;
      A     "B 11.0";
      AN    "M 63.1";
      )     ;
      O     #SERVICE_RUN; // Drive Test - Logic : DON'T CARE!
      A     "M 62.0";
      A     "M 63.0";
      S     "M 63.1";
NETWORK
TITLE =Step 13N3 - Conveyor 12 - Stop Filling

      A     "B 11.0";
      A     "M 62.0";
      A     "M 63.1";
      S     "M 63.2";
NETWORK
TITLE =Step 13N4 - Conveyor 12 - Transfering

      A     "M 67.1";
      AN    "M 67.2";
      A     "M 62.0";
      A     "M 63.2";
      S     "M 63.3";
NETWORK
TITLE =Step 13N5 - Conveyor 12 - Steps Register - Reset

      A(    ;
      O     "B 11.1";
      O     "Timer 63";
      )     ;
      A     "M 62.0";
      A     "M 63.3";
      S     "M 63.4";
NETWORK
TITLE =Conveyor 12 VFD - Release

      A(    ;
      A     "M 63.1";
      AN    "M 63.2";
      O     ;
      A     "M 63.3";
      AN    "M 63.4";
      )     ;
      A     "M 62.0";
      AN    "M 11.1"; // VFD NOT All Ready !
      =     "A 48.6";
      =     "A 48.7";
END_FUNCTION

FUNCTION "NEW C13 - DELIV. LO" : VOID
TITLE =NEW FC966 (was FC1066) - Conveyor 13 - Delivery First Level
NAME : POS_15_L
VERSION : 0.0


VAR_TEMP
  MAIN_SERVICE_2_SW : BOOL ;
  SERVICE_RUN : BOOL ;
  BARRIER_BLINKER : BOOL ;	//Feeder Safety Light Barrier
END_VAR
BEGIN
NETWORK
TITLE =Conveyor 13 - Service

      A     "HMI_DB".ALL_SERVICE_ENABLE_SW;
      A     "HMI_DB".CONVEYOR_11_SERVICE_SW;
      A     "HMI_DB".SERVICE_SW_2_STATUS;
      =     #MAIN_SERVICE_2_SW;
//;
      A     #MAIN_SERVICE_2_SW;
      O     "M 66.1";
      JNB   CO13;
//;
      A     "HMI_DB".HMI_CONVEYOR_13_TEST_SSW;
      =     #SERVICE_RUN;
//;
      AN    #MAIN_SERVICE_2_SW;
      R     "HMI_DB".HMI_CONVEYOR_13_TEST_SSW;

CO13: R     #SERVICE_RUN;
      FP    "FP 148.2";
      =     "M 66.1";
NETWORK
TITLE =Delivery Conveyor 13 - Running TimeOut  30s
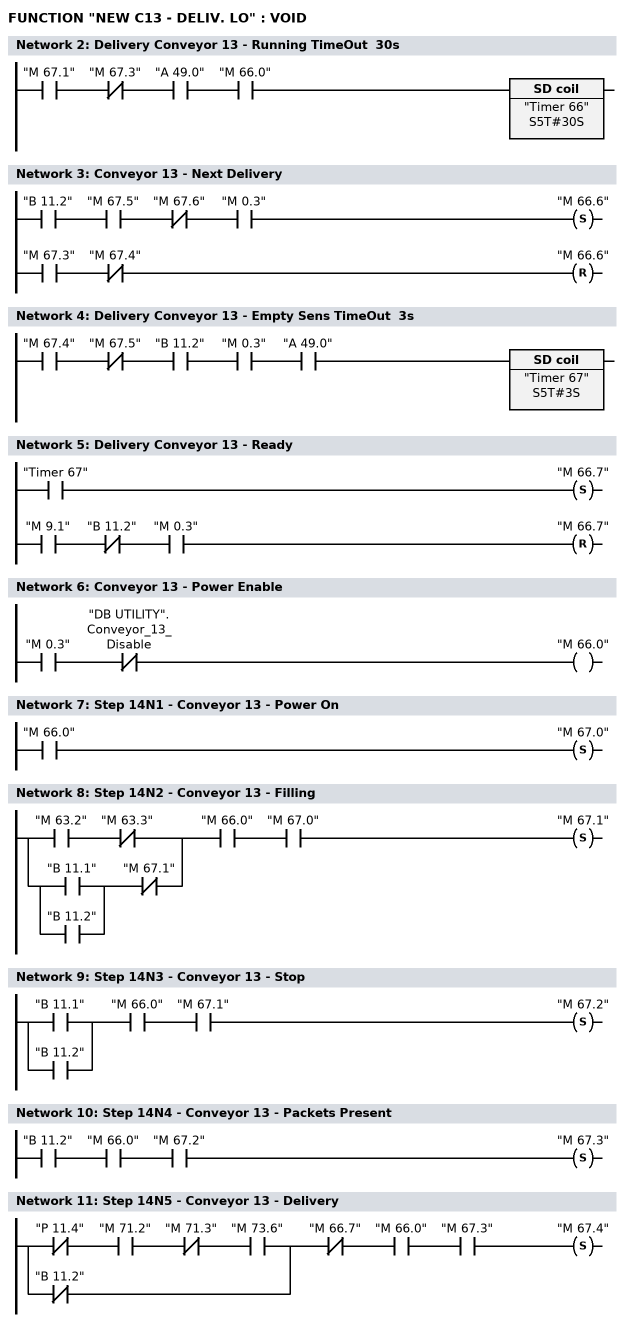

      A     "M 67.1";
      AN    "M 67.3";
      A     "A 49.0";
      A     "M 66.0";
      L     S5T#30S;
      SD    "Timer 66";
NETWORK
TITLE =Conveyor 13 - Next Delivery

      A     "B 11.2";
      A     "M 67.5";
      AN    "M 67.6";
      A     "M 0.3";
      S     "M 66.6";
//;
      A     "M 67.3";
      AN    "M 67.4";
      R     "M 66.6";
NETWORK
TITLE =Delivery Conveyor 13 - Empty Sens TimeOut  3s

      A     "M 67.4";
      AN    "M 67.5";
      A     "B 11.2";
      A     "M 0.3";
      A     "A 49.0";
      L     S5T#3S;
      SD    "Timer 67";
NETWORK
TITLE =Delivery Conveyor 13 - Ready

      A     "Timer 67";
      S     "M 66.7";
//;
      A     "M 9.1";
      AN    "B 11.2";
      A     "M 0.3";
      R     "M 66.7";
NETWORK
TITLE =Conveyor 13 - Power Enable

      A     "M 0.3";
      AN    "DB UTILITY".Conveyor_13_Disable;
      =     "M 66.0";
NETWORK
TITLE =Step 14N1 - Conveyor 13 - Power On

      A     "M 66.0";
      S     "M 67.0";
NETWORK
TITLE =Step 14N2 - Conveyor 13 - Filling

      A(    ;
      A     "M 63.2";
      AN    "M 63.3";
      O     ;
      A(    ;
      O     "B 11.1";
      O     "B 11.2";
      )     ;
//      O     #SERVICE_RUN
      AN    "M 67.1";
      )     ;
      A     "M 66.0";
      A     "M 67.0";
      S     "M 67.1";
NETWORK
TITLE =Step 14N3 - Conveyor 13 - Stop

      A(    ;
      O     "B 11.1";
      O     "B 11.2";
      )     ;
      A     "M 66.0";
      A     "M 67.1";
      S     "M 67.2";
NETWORK
TITLE =Step 14N4 - Conveyor 13 - Packets Present

      A     "B 11.2";
      A     "M 66.0";
      A     "M 67.2";
      S     "M 67.3";
NETWORK
TITLE =Step 14N5 - Conveyor 13 - Delivery

      A(    ;
      AN    "P 11.4";
      A     "M 71.2";
      AN    "M 71.3";
      A     "M 73.6";
      ON    "B 11.2";
      )     ;
      AN    "M 66.7";
      A     "M 66.0";
      A     "M 67.3";
      S     "M 67.4";
NETWORK
TITLE =Write 1 to Steps 0-3 Byte Register MB67

      A(    ;
      O     "M 66.6";
      O     "M 66.7";
      )     ;
      A     "M 67.4";
      A     "M 66.0";
      JC    M001;
      JU    M002;

M001: L     2#1111;
      T     "MB 67";

M002: NOP   0;
NETWORK
TITLE =Step 14N6 - Conveyor 13 - Delivery Done
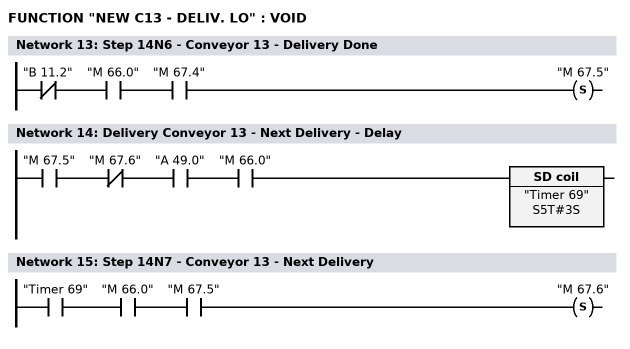

      AN    "B 11.2";
      A     "M 66.0";
      A     "M 67.4";
      S     "M 67.5";
NETWORK
TITLE =Delivery Conveyor 13 - Next Delivery - Delay

      A     "M 67.5";
      AN    "M 67.6";
      A     "A 49.0";
      A     "M 66.0";
      L     S5T#3S;
      SD    "Timer 69";
NETWORK
TITLE =Step 14N7 - Conveyor 13 - Next Delivery

      A     "Timer 69";
      A     "M 66.0";
      A     "M 67.5";
      S     "M 67.6";
NETWORK
TITLE =Steps Register - Reset

      A(    ;
      O     "M 67.6";
      O     "Timer 66";
      )     ;
      A     "M 66.0";
      JC    M003;
      JU    M004;

M003: L     2#0;
      T     "MW 67";

M004: NOP   0;
NETWORK
TITLE =Conveyor 13 VFD - Release
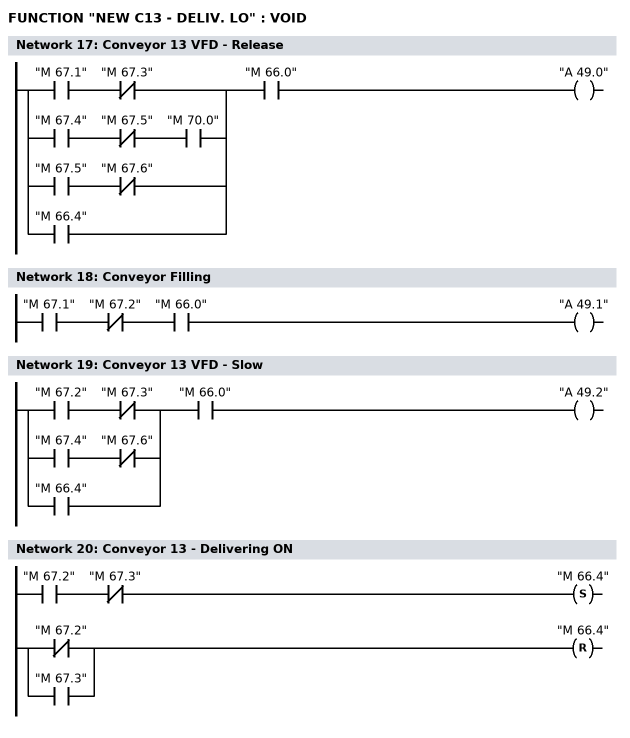

      A(    ;
      A     "M 67.1";
      AN    "M 67.3";
      O     ;
      A     "M 67.4";
      AN    "M 67.5";
      A     "M 70.0";
      O     ;
      A     "M 67.5";
      AN    "M 67.6";
      O     "M 66.4";
      )     ;
      A     "M 66.0";
      =     "A 49.0";
NETWORK
TITLE =Conveyor Filling

      A     "M 67.1";
      AN    "M 67.2";
      A     "M 66.0";
      =     "A 49.1";
NETWORK
TITLE =Conveyor 13 VFD - Slow

      A(    ;
      A     "M 67.2";
      AN    "M 67.3";
      O     ;
      A     "M 67.4";
      AN    "M 67.6";
      O     "M 66.4";
      )     ;
      A     "M 66.0";
      =     "A 49.2";
NETWORK
TITLE =Conveyor 13 - Delivering ON

      A     "M 67.2";
      AN    "M 67.3";
      S     "M 66.4";
//;
      A(    ;
      ON    "M 67.2";
      O     "M 67.3";
      )     ;
      R     "M 66.4";
END_FUNCTION

FUNCTION "NEW LOADER FINGERS" : VOID
TITLE =NEW FC970 (was FC1070) - Feeder Fingers
//
NAME : FEEDER
VERSION : 0.0


VAR_TEMP
  MAIN_SERVICE_3_SW : BOOL ;
  FEEDER_SERVICE_SW : BOOL ;
  FINGERS_SERVICE_SW : BOOL ;
  LIGHT_BARRIER : BOOL ;
  FINGERS_EXTEND : BOOL ;
  FINGERS_RETRACT : BOOL ;
  FINGERS_TILT : BOOL ;
  BELT_ON : BOOL ;
  INITIALISATION : BOOL ;
END_VAR
BEGIN
NETWORK
TITLE =Light Barrier Buffer
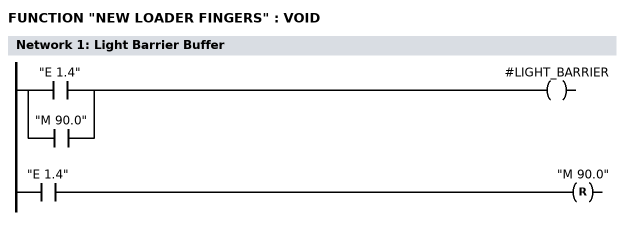

      A     "E 1.4";
      O     "M 90.0";
      =     #LIGHT_BARRIER;
//;
      A     "E 1.4";
      R     "M 90.0";
NETWORK
TITLE =Feeder Service

      A     "HMI_DB".ALL_SERVICE_ENABLE_SW;
      A     "HMI_DB".LOADER_SERVICE_ENABLE_SW;
      A     "HMI_DB".SERVICE_SW_3_STATUS;
      =     #MAIN_SERVICE_3_SW;
//;
      A     #MAIN_SERVICE_3_SW;
      O     "M 70.7";
      JNB   FEED;
      A     "HMI_DB".LOADER_LIFT_SERVICE_SSW;
      =     #FEEDER_SERVICE_SW;
//;
      A     #FEEDER_SERVICE_SW;
      A     "HMI_DB".LOADER_FING_SERVICE_SSW;
      =     #FINGERS_SERVICE_SW;
      =     "DB UTILITY".Conveyor_13_Disable;
      =     "DB UTILITY".Conveyor_23_Disable;
//;
      A     #FEEDER_SERVICE_SW;
      A     #FINGERS_SERVICE_SW;
      A     "HMI_DB".FINGER_EXTEND_TEST_PB;
      AN    #FINGERS_RETRACT;
      =     #FINGERS_EXTEND;
//;
      A     #FEEDER_SERVICE_SW;
      A     #FINGERS_SERVICE_SW;
      A     "HMI_DB".FINGER_RETRACT_TEST_PB;
      AN    #FINGERS_EXTEND;
      =     #FINGERS_RETRACT;
//;
      A     #FEEDER_SERVICE_SW;
      A     #FINGERS_SERVICE_SW;
      A     "HMI_DB".FINGER_BELT_TEST_SW;
      =     #BELT_ON;
//;
      A     #FEEDER_SERVICE_SW;
      A     #FINGERS_SERVICE_SW;
      A     "HMI_DB".FINGER_TILT_TEST_PB;
      =     #FINGERS_TILT;
//;
      AN    #MAIN_SERVICE_3_SW;
      ON    #FEEDER_SERVICE_SW;
      R     "HMI_DB".LOADER_FING_SERVICE_SSW;
      R     "HMI_DB".LOADER_LIFT_SERVICE_SSW;
      R     "HMI_DB".FINGER_RETRACT_TEST_PB;
      R     "HMI_DB".FINGER_EXTEND_TEST_PB;
      R     "HMI_DB".FINGER_TILT_TEST_PB;
      R     "HMI_DB".FINGER_BELT_TEST_SW;

FEED: R     #FEEDER_SERVICE_SW;
      R     #FINGERS_SERVICE_SW;
      R     #FINGERS_EXTEND;
      R     #FINGERS_RETRACT;
      R     #FINGERS_TILT;
      FP    "FP 159.7";
      =     "M 70.7";
//;
      A     "HMI_DB".SERVICE_INIT_PB;
      A     #FEEDER_SERVICE_SW;
      A     #MAIN_SERVICE_3_SW;
      =     #INITIALISATION;
NETWORK
TITLE =Feeder - Power Enable
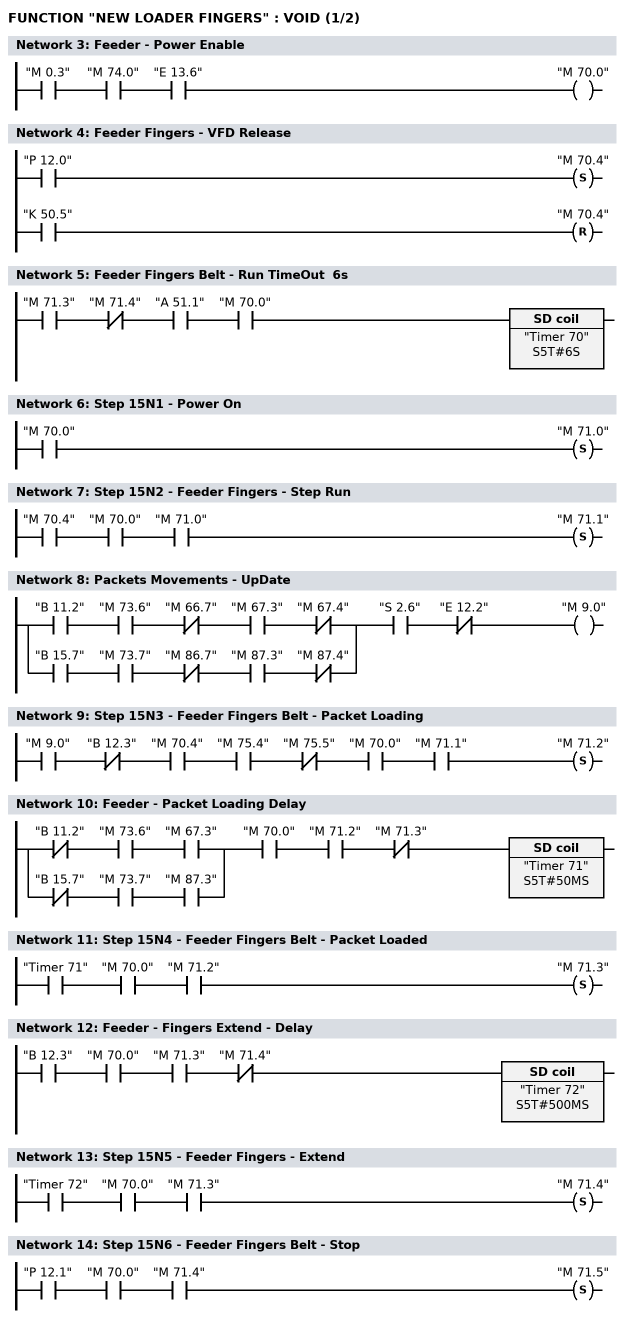

      A     "M 0.3";
      A     "M 74.0";
      A     "E 13.6";
      =     "M 70.0";
NETWORK
TITLE =Feeder Fingers - VFD Release

      A     "P 12.0";
      S     "M 70.4";
//;
      A     "K 50.5";
      R     "M 70.4";
NETWORK
TITLE =Feeder Fingers Belt - Run TimeOut  6s

      A     "M 71.3";
      AN    "M 71.4";
      A     "A 51.1";
      A     "M 70.0";
      L     S5T#6S;
      SD    "Timer 70";
NETWORK
TITLE =Step 15N1 - Power On

      A     "M 70.0";
      S     "M 71.0";
NETWORK
TITLE =Step 15N2 - Feeder Fingers - Step Run

      A     "M 70.4";
      A     "M 70.0";
      A     "M 71.0";
      S     "M 71.1";
NETWORK
TITLE =Packets Movements - UpDate

      A(    ;
      A     "B 11.2";
      A     "M 73.6";
      AN    "M 66.7";
      A     "M 67.3";
      AN    "M 67.4";
      O     ;
      A     "B 15.7";
      A     "M 73.7";
      AN    "M 86.7";
      A     "M 87.3";
      AN    "M 87.4";
      )     ;
      A     "S 2.6";
      AN    "E 12.2";
      =     "M 9.0";
NETWORK
TITLE =Step 15N3 - Feeder Fingers Belt - Packet Loading

      A     "M 9.0";
      AN    "B 12.3";
      A     "M 70.4";
      A     "M 75.4";
      AN    "M 75.5";
      A     "M 70.0";
      A     "M 71.1";
      S     "M 71.2";
NETWORK
TITLE =Feeder - Packet Loading Delay

      A(    ;
      AN    "B 11.2";
      A     "M 73.6";
      A     "M 67.3";
      O     ;
      AN    "B 15.7";
      A     "M 73.7";
      A     "M 87.3";
      )     ;
      A     "M 70.0";
      A     "M 71.2";
      AN    "M 71.3";
      L     S5T#50MS;
      SD    "Timer 71";
NETWORK
TITLE =Step 15N4 - Feeder Fingers Belt - Packet Loaded

      A     "Timer 71";
      A     "M 70.0";
      A     "M 71.2";
      S     "M 71.3";
NETWORK
TITLE =Feeder - Fingers Extend - Delay

      A     "B 12.3";
      A     "M 70.0";
      A     "M 71.3";
      AN    "M 71.4";
      L     S5T#500MS;
      SD    "Timer 72";
NETWORK
TITLE =Step 15N5 - Feeder Fingers - Extend

      A     "Timer 72";
      A     "M 70.0";
      A     "M 71.3";
      S     "M 71.4";
NETWORK
TITLE =Step 15N6 - Feeder Fingers Belt - Stop

      A     "P 12.1";
      A     "M 70.0";
      A     "M 71.4";
      S     "M 71.5";
NETWORK
TITLE =Step 15N7 - Feeder Fingers Tilt - Ready
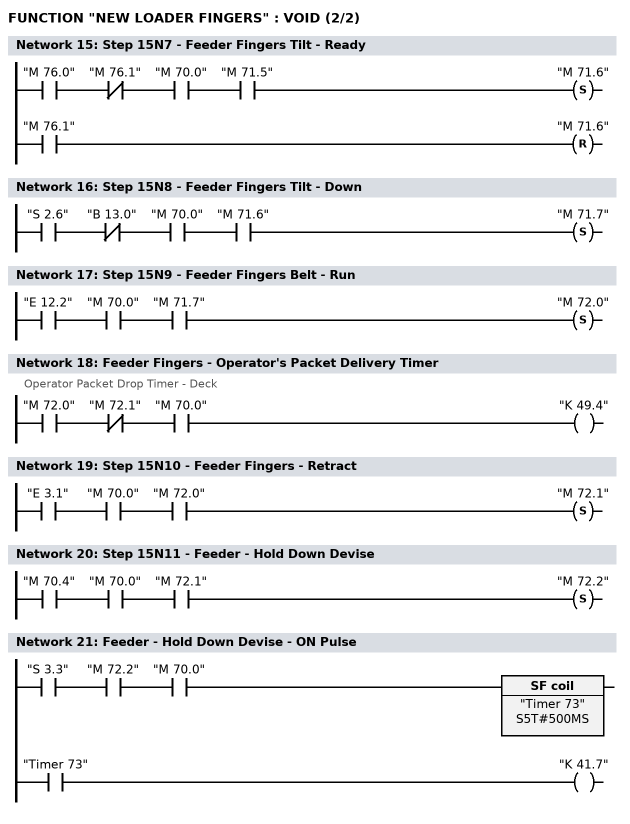

      A     "M 76.0";
      AN    "M 76.1";
      A     "M 70.0";
      A     "M 71.5";
      S     "M 71.6";
//;
      O     "M 76.1";
      R     "M 71.6";
NETWORK
TITLE =Step 15N8 - Feeder Fingers Tilt - Down

      A     "S 2.6";
      AN    "B 13.0";
      A     "M 70.0";
      A     "M 71.6";
      S     "M 71.7";
NETWORK
TITLE =Step 15N9 - Feeder Fingers Belt - Run

      A     "E 12.2";
      A     "M 70.0";
      A     "M 71.7";
      S     "M 72.0";
NETWORK
TITLE =Feeder Fingers - Operator's Packet Delivery Timer
//Operator Packet Drop Timer - Deck
      A     "M 72.0";
      AN    "M 72.1";
      A     "M 70.0";
      =     "K 49.4";
NETWORK
TITLE =Step 15N10 - Feeder Fingers - Retract

      A     "E 3.1";
      A     "M 70.0";
      A     "M 72.0";
      S     "M 72.1";
NETWORK
TITLE =Step 15N11 - Feeder - Hold Down Devise

      A     "M 70.4";
      A     "M 70.0";
      A     "M 72.1";
      S     "M 72.2";
NETWORK
TITLE =Feeder - Hold Down Devise - ON Pulse

      A     "S 3.3";
      A     "M 72.2";
      A     "M 70.0";
      L     S5T#500MS;
      SF    "Timer 73";

      A     "Timer 73";
      =     "K 41.7";
NETWORK
TITLE =Feeder Fingers - Steps Chain Register Reset

      A(    ;
      ON    "M 75.0";
      O     "M 72.2";
      O     "Timer 70";
      O     #FEEDER_SERVICE_SW;
      )     ;
      JC    M001;
      JU    M002;

M001: L     2#0;
      T     "MW 71";

M002: NOP   0;
NETWORK
TITLE =Feeder Fingers - Fingers Retract
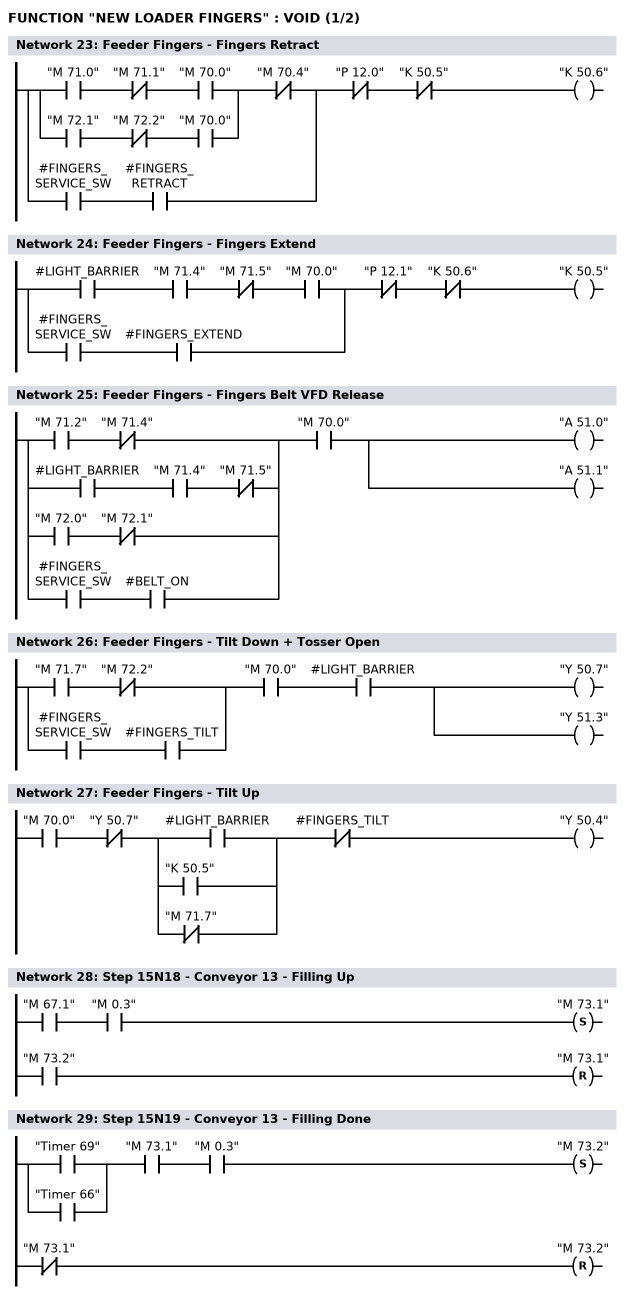

      A(    ;
      A(    ;
      A     "M 71.0";
      AN    "M 71.1";
      A     "M 70.0";
      O     ;
      A     "M 72.1";
      AN    "M 72.2";
      A     "M 70.0";
      )     ;
      AN    "M 70.4";
      O     ;
      A     #FINGERS_SERVICE_SW;
      A     #FINGERS_RETRACT;
      )     ;
      AN    "P 12.0";
      AN    "K 50.5";
      =     "K 50.6";
NETWORK
TITLE =Feeder Fingers - Fingers Extend

      A(    ;
      A     #LIGHT_BARRIER;
      A     "M 71.4";
      AN    "M 71.5";
      A     "M 70.0";
      O     ;
      A     #FINGERS_SERVICE_SW;
      A     #FINGERS_EXTEND;
      )     ;
      AN    "P 12.1";
      AN    "K 50.6";
      =     "K 50.5";
NETWORK
TITLE =Feeder Fingers - Fingers Belt VFD Release

      A(    ;
      A     "M 71.2";
      AN    "M 71.4";
      O     ;
      A     #LIGHT_BARRIER;
      A     "M 71.4";
      AN    "M 71.5";
      O     ;
      A     "M 72.0";
      AN    "M 72.1";
      O     ;
      A     #FINGERS_SERVICE_SW;
      A     #BELT_ON;
      )     ;
      A     "M 70.0";
      =     "A 51.0";
      =     "A 51.1";
NETWORK
TITLE =Feeder Fingers - Tilt Down + Tosser Open

      A(    ;
      A     "M 71.7";
      AN    "M 72.2";
      O     ;
      A     #FINGERS_SERVICE_SW;
      A     #FINGERS_TILT;
      )     ;
      A     "M 70.0";
      A     #LIGHT_BARRIER;
      =     "Y 50.7";
      =     "Y 51.3";
NETWORK
TITLE =Feeder Fingers - Tilt Up

      A     "M 70.0";
      AN    "Y 50.7";
      A(    ;
      O     #LIGHT_BARRIER;
      O     "K 50.5";
      ON    "M 71.7";
      AN    #FINGERS_TILT;
      )     ;
      =     "Y 50.4";
NETWORK
TITLE =Step 15N18 - Conveyor 13 - Filling Up

      A     "M 67.1";
      A     "M 0.3";
      S     "M 73.1";
//;
      A     "M 73.2";
      R     "M 73.1";
NETWORK
TITLE =Step 15N19 - Conveyor 13 - Filling Done

      A(    ;
      O     "Timer 69";
      O     "Timer 66";
      )     ;
      A     "M 73.1";
      A     "M 0.3";
      S     "M 73.2";
//;
      AN    "M 73.1";
      R     "M 73.2";
NETWORK
TITLE =Step 15N20 - Conveyor 23 - Filling Up
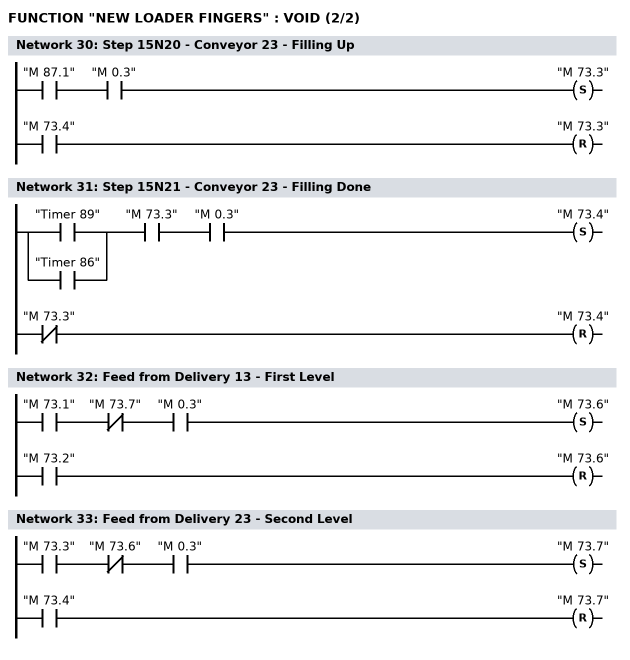

      A     "M 87.1";
      A     "M 0.3";
      S     "M 73.3";
//;
      A     "M 73.4";
      R     "M 73.3";
NETWORK
TITLE =Step 15N21 - Conveyor 23 - Filling Done

      A(    ;
      O     "Timer 89";
      O     "Timer 86";
      )     ;
      A     "M 73.3";
      A     "M 0.3";
      S     "M 73.4";
//;
      AN    "M 73.3";
      R     "M 73.4";
NETWORK
TITLE =Feed from Delivery 13 - First Level

      A     "M 73.1";
      AN    "M 73.7";
      A     "M 0.3";
      S     "M 73.6";
//;
      A     "M 73.2";
      R     "M 73.6";
NETWORK
TITLE =Feed from Delivery 23 - Second Level

      A     "M 73.3";
      AN    "M 73.6";
      A     "M 0.3";
      S     "M 73.7";
//;
      A     "M 73.4";
      R     "M 73.7";
END_FUNCTION

FUNCTION "NEW LOADER LIFT" : VOID
TITLE =NEW FC974 (was FC1074) - Feeder Lift Pos. 16
//
NAME : FEEDER
VERSION : 0.0


VAR_TEMP
  MAIN_SERVICE_3_SW : BOOL ;
  FEEDER_SW : BOOL ;
  FEEDER_SERVICE_SW : BOOL ;
  LIGHT_BARRIER : BOOL ;
  FEEDER_LIFT_TOP_PB : BOOL ;
  FEEDER_LIFT_UP_PB : BOOL ;
  FEEDER_LIFT_DN_PB : BOOL ;
  FEEDER_LIFT_JOG_UP : BOOL ;
  FEEDER_LIFT_JOG_DN : BOOL ;
END_VAR
BEGIN
NETWORK
TITLE =Light Barrier Buffer
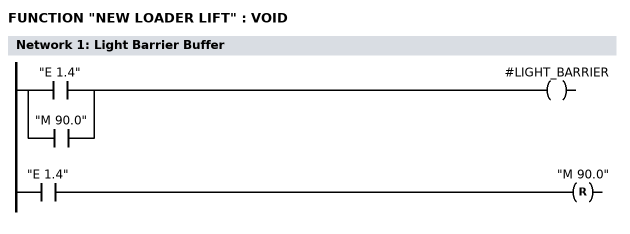

      A     "E 1.4";
      O     "M 90.0";
      =     #LIGHT_BARRIER;
//;
      A     "E 1.4";
      R     "M 90.0";
NETWORK
TITLE =Feeder Service

      A     "HMI_DB".ALL_SERVICE_ENABLE_SW;
      A     "HMI_DB".LOADER_SERVICE_ENABLE_SW;
      A     "HMI_DB".SERVICE_SW_3_STATUS;
      =     #MAIN_SERVICE_3_SW;
//;
      A     #MAIN_SERVICE_3_SW;
      O     "M 74.7";
      JNB   FEED;
      A     "HMI_DB".LOADER_LIFT_SERVICE_SSW;
      =     #FEEDER_SERVICE_SW;
      S     "DB UTILITY".Conveyor_13_Disable;
      S     "DB UTILITY".Conveyor_23_Disable;
      R     "M 74.2";
//;
      A     #FEEDER_SERVICE_SW;
      A     "HMI_DB".LOADER_LIFT_TOP_PB;
      =     #FEEDER_LIFT_TOP_PB;
//;
      A     #FEEDER_SERVICE_SW;
      A     "HMI_DB".LOADER_LIFT_UP_PB;
      =     #FEEDER_LIFT_UP_PB;
//;
      A     #FEEDER_SERVICE_SW;
      A     "HMI_DB".LOADER_LIFT_DN_PB;
      =     #FEEDER_LIFT_DN_PB;
//;
      AN    #MAIN_SERVICE_3_SW;
      ON    #FEEDER_SERVICE_SW;
      R     "HMI_DB".LOADER_FING_SERVICE_SSW;
      R     "HMI_DB".LOADER_LIFT_SERVICE_SSW;
      R     "HMI_DB".LOADER_LIFT_TOP_PB;
      R     "HMI_DB".LOADER_LIFT_UP_PB;
      R     "HMI_DB".LOADER_LIFT_DN_PB;
      R     "DB UTILITY".Conveyor_13_Disable;
      R     "DB UTILITY".Conveyor_23_Disable;

FEED: R     #FEEDER_SERVICE_SW;
      R     #FEEDER_LIFT_TOP_PB;
      R     #FEEDER_LIFT_UP_PB;
      R     #FEEDER_LIFT_DN_PB;
      FP    "FP 159.6";
      =     "M 74.7";
NETWORK
TITLE =Automatic Trigger
